(* IEC 61131-3 sources: plcassist-cli/packages/volt-lsp-iec/test-corpus/lenze-mid/Device/Plc Logic/Application/Library Manager/L_MC4P_RoboticHandling (part 2) *)

(* ---- L_MC4P_GROUPDIGITALSWITCHHANDLER.fb ---- *)
FUNCTION_BLOCK L_MC4P_GROUPDIGITALSWITCHHANDLER EXTENDS L_MC4P_Template_AG_KIN
VAR_INPUT
	XENABLE : BOOL;
	XRESETSWITCHES : BOOL;
END_VAR
VAR_OUTPUT
	XVALID : BOOL;
	XBUSY : BOOL;
	XERROR : BOOL;
	EERRORID : L_IE1P_Error;
	DWDIGITALSWITCHES : DWORD;
END_VAR
VAR
	ADWDIGITALSWITCHES : ARRAY [1..cwNbrOfdwDigSwitches] OF DWORD;
	LRPASSEDLENGTHOFSEGMENTID : LREAL;
	LRPASSEDTIMEOFSEGMENTID : LREAL;
	_MODEL : L_UBUP_BehaviourModel_LCon;
	XRESETSWITCHESOLD : BOOL;
	RSCSWITCHINGFUN : REFERENCE TO L_MC4P_SwitchingFunctionData;
	ALRSWITCHPARAMSORTED : ARRAY [1..L_MC4P_Constants.gciMaxNumParallelSwitchingFun] OF LREAL;
	XPOSRELATED : BOOL;
	ISWITCHIDXVISU : INT := 1;
	WVISUIDX : WORD := 1;
	CWNBROFDWDIGSWITCHES : WORD := 1024;
	IDXMAX : DINT;
	IDXMIN : DINT;
END_VAR
END_FUNCTION_BLOCK

METHOD ANALYZEANDSORTDATA : BOOL
VAR_INPUT
	PLISTELEMENT : POINTER TO L_MC4P_ListElement;
END_VAR
END_METHOD

METHOD GETDIGITALSWITCH : BOOL
VAR_INPUT
	WDIGITALSWITCH : WORD;
END_VAR
END_METHOD

METHOD RESET : BOOL
END_METHOD

METHOD SETDIGITALSWITCH : BOOL
VAR_INPUT
	WDIGITALSWITCH : WORD;
	XVALUE : BOOL;
END_VAR
END_METHOD

METHOD SETEVALUATEDFLAG : BOOL
VAR_INPUT
	PLISTELEMENT : POINTER TO L_MC4P_ListElement;
	IDX : INT;
END_VAR
END_METHOD

METHOD SPLITINDEX : BOOL
VAR_INPUT
	WSWITCHIDX : WORD;
END_VAR
VAR_OUTPUT
	WARRIDX : WORD;
	WBITIDX : WORD;
END_VAR
END_METHOD

METHOD CYCLICIPOCALL : BOOL
VAR_INPUT
	PLISTELEMENT : POINTER TO L_MC4P_ListElement;
	RSCCYCLICDATA : REFERENCE TO L_MC4P_CyclicData;
END_VAR
END_METHOD

METHOD FINALIZESEGMENT : BOOL
VAR_INPUT
	PLISTELEMENTACT : POINTER TO L_MC4P_ListElement;
	PLISTELEMENTNEXT : POINTER TO L_MC4P_ListElement;
END_VAR
END_METHOD

METHOD CYCLICACTION
VAR_INPUT
	ITFTIMINGCONTROLLER : L_UBUP.L_UBUP_ITimingController;
END_VAR
VAR_OUTPUT
	XCOMPLETE : BOOL;
	XABORT : BOOL;
	IERRORID : INT;
END_VAR
END_METHOD

METHOD FINALIZEACTION
VAR_INPUT
	XABORTPROPOSED : BOOL;
	IERRORIDPROPOSED : INT;
END_VAR
VAR_OUTPUT
	XCOMPLETE : BOOL;
	XABORT : BOOL;
	IERRORID : INT;
END_VAR
END_METHOD

METHOD RESETACTION
VAR_OUTPUT
	XCOMPLETE : BOOL;
END_VAR
END_METHOD

METHOD STARTACTION
VAR_OUTPUT
	XCOMPLETE : BOOL;
	IERRORID : INT;
END_VAR
END_METHOD

METHOD EXCHANGE : BOOL
VAR_INPUT
	IDX1 : DINT;
	IDX2 : DINT;
END_VAR
END_METHOD

METHOD GETVALUE : LREAL
VAR_INPUT
	IDX : DINT;
END_VAR
END_METHOD

(* ---- L_MC4P_GROUPHOME_INTERNAL.fb ---- *)
FUNCTION_BLOCK L_MC4P_GROUPHOME_INTERNAL EXTENDS L_UBUP_PoolInstance
VAR_INPUT
	EXECUTE : BOOL;
END_VAR
VAR_OUTPUT
	DONE : BOOL;
	BUSY : BOOL;
	ACTIVE : BOOL;
	COMMANDABORTED : BOOL;
	ERROR : BOOL;
	ERRORID : L_IE1P_Error;
	AXISDONE : ARRAY [1..12] OF BOOL;
END_VAR
VAR
	COORDSYSTEM : L_MC4P_CoordSystem := L_MC4P_CoordSystem.ACS;
	AMC_HOME : ARRAY [1..12] OF L_MC1P_Home_Internal;
	AMC_HOME_FBBASE : ARRAY [1..12] OF L_MC1P_Template;
	XRESETOUTPUT : BOOL;
	XEXECUTEOLD : BOOL;
	XVALIDAXISSTATES : BOOL;
	IDX : WORD;
	EACTHOMINGORDER : L_MC4P_HomingOrder := L_MC4P_HomingOrder.NoHoming;
	AXAXESHOMED : ARRAY [1..12] OF BOOL;
	ALRPOSITION_INT : ARRAY [1..12] OF LREAL;
	AEHOMINGORDER_INT : ARRAY [1..12] OF L_MC4P_HomingOrder := [12(0)];
	ECOORDSYSTEM_INT : L_MC4P_CoordSystem;
	ASCEXTPARAMETER_INT : ARRAY [1..12] OF L_MC1P_HomeParameter;
	AXUSEEXTPARAMETER_INT : ARRAY [1..12] OF BOOL;
	ASCEXTTP_INT : ARRAY [1..12] OF MC_TRIGGER_REF;
	CLASSID : DINT;
END_VAR
END_FUNCTION_BLOCK

METHOD MAIN
VAR_IN_OUT
	AXESGROUP : AXES_GROUP_KIN;
	FBBASE : L_MC4P_Template_AG_KIN;
	POSITION : ARRAY [1..12] OF LREAL;
	HOMINGORDER : ARRAY [1..12] OF L_MC4P_HomingOrder;
	HOMEABSSWITCH : ARRAY [1..12] OF BOOL;
	USEEXTPARAMETER : ARRAY [1..12] OF BOOL;
	EXTPARAMETER : ARRAY [1..12] OF L_MC1P_HomeParameter;
	EXTTP : ARRAY [1..12] OF MC_TRIGGER_REF;
END_VAR
END_METHOD

METHOD RESETOUTPUTS
END_METHOD

METHOD SETAXISMC_HOME_ACS : BOOL
VAR_IN_OUT
	AXESGROUP : AXES_GROUP_KIN;
	FBBASE : L_MC4P_Template_AG_KIN;
	HOMEABSSWITCH : ARRAY [1..12] OF BOOL;
END_VAR
END_METHOD

METHOD SETNEXTHOMESTEP
END_METHOD

METHOD GET_EERRORID : L_IE1P_Error
END_METHOD

METHOD GET_XACTIVE : BOOL
END_METHOD

METHOD GET_XBUSY : BOOL
END_METHOD

METHOD GET_XCOMMANDABORTED : BOOL
END_METHOD

METHOD GET_XDONE : BOOL
END_METHOD

METHOD GET_XINITIAL : BOOL
END_METHOD

METHOD FREE : BOOL
END_METHOD

(* ---- L_MC4P_GROUPMANUALMODE.fb ---- *)
FUNCTION_BLOCK L_MC4P_GROUPMANUALMODE EXTENDS L_MC4P_Template_AG_KIN
VAR_INPUT
	ALRSETPOSDIST : ARRAY [1..12] OF LREAL;
	SCPAR : L_MC4P_GroupManualMode_Parameter;
	ECOORDSYSTEM : L_MC4P_CoordSystem;
	AXJOGPOS : ARRAY [1..12] OF BOOL;
	AXJOGNEG : ARRAY [1..12] OF BOOL;
	AXMOVEABSEXECUTE : ARRAY [1..12] OF BOOL;
	AXMOVERELEXECUTE : ARRAY [1..12] OF BOOL;
END_VAR
VAR_OUTPUT
	XINTERNALCONTROLACTIVE : BOOL;
	XBUSY : BOOL;
	XDONE : BOOL;
	XERROR : BOOL;
	EERRORID : L_IE1P_Error;
	EMANUALMODE : L_MC4P_ManualMode := L_MC4P_ManualMode.Standby;
END_VAR
VAR
	MANMODE : L_MC4P_GroupManualMode_Internal;
END_VAR
END_FUNCTION_BLOCK

(* ---- L_MC4P_GROUPMANUALMODE_INTERNAL.fb ---- *)
FUNCTION_BLOCK L_MC4P_GROUPMANUALMODE_INTERNAL EXTENDS L_UBUP_PoolInstance
VAR_INPUT
	ALRSETPOSDIST : ARRAY [1..12] OF LREAL;
	SCPAR : L_MC4P_GroupManualMode_Parameter;
	ECOORDSYSTEM : L_MC4P_CoordSystem;
	AXJOGPOS : ARRAY [1..12] OF BOOL;
	AXJOGNEG : ARRAY [1..12] OF BOOL;
	AXMOVEABSEXECUTE : ARRAY [1..12] OF BOOL;
	AXMOVERELEXECUTE : ARRAY [1..12] OF BOOL;
	XISV2 : BOOL := FALSE;
END_VAR
VAR_OUTPUT
	XINTERNALCONTROLACTIVE : BOOL;
	XBUSY : BOOL;
	XDONE : BOOL;
	XERROR : BOOL;
	EERRORID : L_IE1P_Error;
	EMANUALMODE : L_MC4P_ManualMode := L_MC4P_ManualMode.Standby;
END_VAR
VAR
	AXMOVEABSEXECUTEEDGE : ARRAY [1..12] OF BOOL;
	AXMOVERELEXECUTEEDGE : ARRAY [1..12] OF BOOL;
	ECOORDSYSTEM_INT : L_MC4P_CoordSystem := L_MC4P_CoordSystem.MCS;
	XDOSTATEMACHINE : BOOL;
	XCHANGETOSTANDBY : BOOL := FALSE;
	XJOGGING : BOOL;
	XMOVEABSEDGE : BOOL;
	XMOVERELEDGE : BOOL;
	XMOVEABS : BOOL;
	XMOVEREL : BOOL;
	AMANUALJOG : ARRAY [1..12] OF L_MC1P_ManualJog_Internal;
	AMANUALJOG_FBBASE : ARRAY [1..12] OF L_MC1P.L_MC1P_Template;
	AMC_MOVERELATIVE : ARRAY [1..12] OF L_MC1P_MoveRelative_Internal;
	AMC_MOVERELATIVE_FBBASE : ARRAY [1..12] OF L_MC1P.L_MC1P_Template;
	AMC_MOVEABSOLUTE : ARRAY [1..12] OF L_MC1P_MoveAbsolute_Inernal;
	AMC_MOVEABSOLUTE_FBBASE : ARRAY [1..12] OF L_MC1P.L_MC1P_Template;
	EMANUALMODEOLD : L_MC4P_ManualMode := L_MC4P_ManualMode.Standby;
	ECOORDSYSTEMOLD : L_MC4P_CoordSystem;
	AXMOVEABSEXECUTEOLD : ARRAY [1..12] OF BOOL;
	AXMOVERELEXECUTEOLD : ARRAY [1..12] OF BOOL;
	XMOTIONACTIVE : BOOL := FALSE;
	APG : ARRAY [1..6] OF L_MC1P.L_MC1P_PosProfiler;
	ASCPROFILEPARAMETER : ARRAY [1..6] OF L_MC1P_ProfileParameter;
	PCOORDTRAFO : POINTER TO L_MC4P_CoordTrafo;
	COORDTRAFO_INT : L_MC4P_CoordTrafo;
	ALRPCSSETPOSATEXECUTE : ARRAY [1..6] OF LREAL;
	PLRDUMMY : POINTER TO LREAL;
	ALRPCSSETPOS_EXT : ARRAY [1..6] OF LREAL;
	ALRWCSSETPOS_EXT : ARRAY [1..6] OF LREAL;
	CLASSID : DINT;
END_VAR
END_FUNCTION_BLOCK

METHOD MAIN
VAR_IN_OUT
	AXESGROUP : AXES_GROUP_KIN;
	FBBASE : L_MC4P_Template_AG_KIN;
END_VAR
END_METHOD

METHOD GET_EERRORID : L_IE1P_Error
END_METHOD

METHOD GET_XACTIVE : BOOL
END_METHOD

METHOD GET_XBUSY : BOOL
END_METHOD

METHOD GET_XCOMMANDABORTED : BOOL
END_METHOD

METHOD GET_XDONE : BOOL
END_METHOD

METHOD GET_XINITIAL : BOOL
END_METHOD

METHOD FREE : BOOL
END_METHOD

METHOD CHECKPCSMCS : BOOL
END_METHOD

METHOD ENTRYSTANDBYSTATE
VAR_IN_OUT
	AXESGROUP : AXES_GROUP_KIN;
	FBBASE : L_MC4P_Template_AG_KIN;
END_VAR
END_METHOD

METHOD EXITMOVESTATE
VAR_IN_OUT
	AXESGROUP : AXES_GROUP_KIN;
	FBBASE : L_MC4P_Template_AG_KIN;
END_VAR
END_METHOD

METHOD GETTCSPOSINPCSMCS
VAR_INPUT
	EROTATIONCONVENTIONPCS : L_UMTP_RotationConvention;
END_VAR
VAR_IN_OUT
	AXESGROUP : AXES_GROUP_KIN;
	ALRPCSSETPOS : ARRAY [1..6] OF LREAL;
END_VAR
END_METHOD

METHOD ISMOTIONALLOWED
VAR_IN_OUT
	AXESGROUP : AXES_GROUP_KIN;
	FBBASE : L_MC4P_Template_AG_KIN;
	SCPAR : L_MC4P_GroupManualMode_Parameter;
	ECOORDSYSTEM : L_MC4P_CoordSystem;
	AXJOGPOS : ARRAY [1..12] OF BOOL;
	AXJOGNEG : ARRAY [1..12] OF BOOL;
	AXMOVEABSEXECUTE : ARRAY [1..12] OF BOOL;
	AXMOVERELEXECUTE : ARRAY [1..12] OF BOOL;
END_VAR
END_METHOD

METHOD JOGAXISREF
VAR_INPUT
	XWCS : BOOL;
	XACS : BOOL;
	XAUX : BOOL;
END_VAR
VAR_IN_OUT
	AXESGROUP : AXES_GROUP_KIN;
	FBBASE : L_MC4P_Template_AG_KIN;
	SCPAR : L_MC4P_GroupManualMode_Parameter;
	AXJOGPOS : ARRAY [1..12] OF BOOL;
	AXJOGNEG : ARRAY [1..12] OF BOOL;
END_VAR
END_METHOD

METHOD JOGPCSMCS
VAR_IN_OUT
	AXESGROUP : AXES_GROUP_KIN;
	FBBASE : L_MC4P_Template_AG_KIN;
	SCPAR : L_MC4P_GroupManualMode_Parameter;
	AXJOGPOS : ARRAY [1..12] OF BOOL;
	AXJOGNEG : ARRAY [1..12] OF BOOL;
END_VAR
END_METHOD

METHOD MOVEABSAXISREF
VAR_INPUT
	XWCS : BOOL;
	XACS : BOOL;
	XAUX : BOOL;
END_VAR
VAR_IN_OUT
	AXESGROUP : AXES_GROUP_KIN;
	FBBASE : L_MC4P_Template_AG_KIN;
	ALRSETPOSDIST : ARRAY [1..12] OF LREAL;
	SCPAR : L_MC4P_GroupManualMode_Parameter;
	AXMOVEABSEXECUTE : ARRAY [1..12] OF BOOL;
END_VAR
END_METHOD

METHOD MOVEABSPCSMCS
VAR_IN_OUT
	AXESGROUP : AXES_GROUP_KIN;
	FBBASE : L_MC4P_Template_AG_KIN;
	ALRSETPOSDIST : ARRAY [1..12] OF LREAL;
	SCPAR : L_MC4P_GroupManualMode_Parameter;
	AXMOVEABSEXECUTE : ARRAY [1..12] OF BOOL;
END_VAR
END_METHOD

METHOD MOVERELAXISREF
VAR_INPUT
	XWCS : BOOL;
	XACS : BOOL;
	XAUX : BOOL;
END_VAR
VAR_IN_OUT
	AXESGROUP : AXES_GROUP_KIN;
	FBBASE : L_MC4P_Template_AG_KIN;
	ALRSETPOSDIST : ARRAY [1..12] OF LREAL;
	SCPAR : L_MC4P_GroupManualMode_Parameter;
	AXMOVERELEXECUTE : ARRAY [1..12] OF BOOL;
END_VAR
END_METHOD

METHOD MOVERELPCSMCS
VAR_IN_OUT
	AXESGROUP : AXES_GROUP_KIN;
	FBBASE : L_MC4P_Template_AG_KIN;
	ALRSETPOSDIST : ARRAY [1..12] OF LREAL;
	SCPAR : L_MC4P_GroupManualMode_Parameter;
	AXMOVERELEXECUTE : ARRAY [1..12] OF BOOL;
END_VAR
END_METHOD

METHOD RESETMOTIONQUERY
END_METHOD

METHOD WRITEPCSMCSPOS2AXES
VAR_INPUT
	EROTATIONCONVENTIONPCS : L_UMTP_RotationConvention;
	XRELATIVE : BOOL;
END_VAR
VAR_IN_OUT
	AXESGROUP : AXES_GROUP_KIN;
	FBBASE : L_MC4P_Template_AG_KIN;
	ALRPCSSETPOS : ARRAY [1..6] OF LREAL;
	ALRPCSSETVEL : ARRAY [1..6] OF LREAL;
END_VAR
END_METHOD

METHOD CALL_AXISREFPARM
VAR_INPUT
	AXESGROUP : REFERENCE TO AXES_GROUP_KIN;
	LRVELOCITY : REFERENCE TO LREAL;
	LRACCELERATION : REFERENCE TO LREAL;
	LRDECELERATION : REFERENCE TO LREAL;
	LRJERK : REFERENCE TO LREAL;
	AXIS_IDX_LOCAL : WORD;
END_VAR
END_METHOD

METHOD CALL_PCSMCSPARM
VAR_INPUT
	AXESGROUP : REFERENCE TO AXES_GROUP_KIN;
	ALRPCSSETPOS : REFERENCE TO ARRAY [1..6] OF LREAL;
	IDX_LOCAL : WORD;
END_VAR
END_METHOD

(* ---- L_MC4P_GROUPPOWER.fb ---- *)
FUNCTION_BLOCK L_MC4P_GROUPPOWER EXTENDS L_MC4P_Template_AG_REF
VAR_INPUT
	XENABLE : BOOL;
	AEAXISENABLE : ARRAY [1..12] OF L_MC4P_AxisEnableMode := [12(L_MC4P_AxisEnableMode.EnablePosNeg)];
END_VAR
VAR_OUTPUT
	XSTATUS : BOOL;
	XVALID : BOOL;
	XERROR : BOOL;
	EERRORID : L_IE1P_Error;
END_VAR
VAR
	AMC_POWER : ARRAY [1..12] OF MC_Power;
	XENABLEOLD : BOOL;
	IDX : WORD;
	IDX_PLUSSIX : WORD;
	XAXISEXTENABLED : BOOL := FALSE;
	XERRORINTERN : BOOL := FALSE;
	EERRORIDINTERN : L_IE1P_Error;
	XAXISERROR : BOOL := FALSE;
END_VAR
END_FUNCTION_BLOCK

(* ---- L_MC4P_GROUPREADACTUALPOSITION_INTERNAL.fb ---- *)
FUNCTION_BLOCK L_MC4P_GROUPREADACTUALPOSITION_INTERNAL EXTENDS L_UBUP_Instance
VAR_INPUT
	ENABLE : BOOL;
	COORDSYSTEM : L_MC4P_CoordSystem;
END_VAR
VAR_OUTPUT
	VALID : BOOL;
	BUSY : BOOL;
	ERROR : BOOL;
	ERRORID : L_IE1P_Error;
END_VAR
VAR
	IDX : WORD;
	XENABLEOLD : BOOL;
	PCOORDTRAFO : POINTER TO L_MC4P_CoordTrafo;
	ALRPOSITIONTMP : ARRAY [1..6] OF LREAL;
	CLASSID : DINT;
END_VAR
END_FUNCTION_BLOCK

METHOD MAIN
VAR_INPUT
	XUSESETVALUES : BOOL;
END_VAR
VAR_IN_OUT
	AXESGROUP : AXES_GROUP_KIN;
	FBBASE : L_MC4P_Template_AG_KIN;
	POSITION : ARRAY [1..12] OF LREAL;
END_VAR
END_METHOD

(* ---- L_MC4P_GROUPREADACTUALVELOCITY_INTERNAL.fb ---- *)
FUNCTION_BLOCK L_MC4P_GROUPREADACTUALVELOCITY_INTERNAL EXTENDS L_UBUP_Instance
VAR_INPUT
	ENABLE : BOOL;
	COORDSYSTEM : L_MC4P_CoordSystem;
END_VAR
VAR_OUTPUT
	VALID : BOOL;
	BUSY : BOOL;
	ERROR : BOOL;
	ERRORID : L_IE1P_Error;
END_VAR
VAR
	IDX : WORD;
	XENABLEOLD : BOOL;
	ALRVELOCITYTMP1 : ARRAY [1..6] OF LREAL;
	ALRVELOCITYTMP2 : ARRAY [1..6] OF LREAL;
	ALRPOSITIONTMP : ARRAY [1..6] OF LREAL;
	PCOORDTRAFO : POINTER TO L_MC4P_CoordTrafo;
	ALRPOSVEKPCS2TCS : ARRAY [1..3] OF LREAL;
	ROT_MAT : ARRAY [1..3, 1..3] OF LREAL;
	T4 : LREAL;
	T5 : LREAL;
	T7 : LREAL;
	CLASSID : DINT;
END_VAR
END_FUNCTION_BLOCK

METHOD MAIN
VAR_INPUT
	XUSESETVALUES : BOOL;
END_VAR
VAR_IN_OUT
	AXESGROUP : AXES_GROUP_KIN;
	FBBASE : L_MC4P_Template_AG_KIN;
	VELOCITY : ARRAY [1..12] OF LREAL;
	PATHVELOCITY : LREAL;
END_VAR
END_METHOD

(* ---- L_MC4P_GROUPREADSTATUS_INTERNAL.fb ---- *)
FUNCTION_BLOCK L_MC4P_GROUPREADSTATUS_INTERNAL EXTENDS L_UBUP_PoolInstance
VAR_INPUT
	ENABLE : BOOL;
END_VAR
VAR_OUTPUT
	VALID : BOOL;
	BUSY : BOOL;
	ERROR : BOOL;
	ERRORID : L_IE1P_Error;
	GROUPMOVING : BOOL;
	GROUPHOMING : BOOL;
	GROUPERRORSTOP : BOOL;
	GROUPSTANDBY : BOOL;
	GROUPSTOPPING : BOOL;
	GROUPDISABLED : BOOL;
	CONSTANTVELOCITY : BOOL;
	ACCELERATING : BOOL;
	DECELERATING : BOOL;
	INPOSITION : BOOL;
	STANDSTILL : BOOL;
END_VAR
VAR
	XENABLEOLD : BOOL;
	IDX : INT;
	CLASSID : DINT;
END_VAR
END_FUNCTION_BLOCK

METHOD MAIN
VAR_IN_OUT
	AXESGROUP : AXES_GROUP_KIN;
	FBBASE : L_MC4P_Template_AG_KIN;
END_VAR
END_METHOD

(* ---- L_MC4P_GROUPRESET_INTERNAL.fb ---- *)
FUNCTION_BLOCK L_MC4P_GROUPRESET_INTERNAL EXTENDS L_UBUP_Instance
VAR_INPUT
	EXECUTE : BOOL;
END_VAR
VAR_OUTPUT
	DONE : BOOL;
	BUSY : BOOL;
	ERROR : BOOL;
	ERRORID : L_IE1P_Error;
END_VAR
VAR
	ARESET : ARRAY [1..18] OF MC_Reset;
	PAXESGROUP : POINTER TO AXES_GROUP_KIN;
	XEXECUTEOLD : BOOL;
	PWTMP : POINTER TO WORD;
	IDX : INT;
	XRESETPOSSIBLE : BOOL;
	XRESETOUTPUT : BOOL;
	DWRESETCYCLECOUNTERSTART : DWORD;
	XNOERRORACTIVE : BOOL;
	XERRORSTOPDONE : BOOL;
	XAXESGROUPINERROR : BOOL;
	XAXISINERROR : BOOL;
	XWAITFORRESETEVENT : BOOL;
	DWMAXTIMEOUT : DWORD;
	CLASSID : DINT;
END_VAR
END_FUNCTION_BLOCK

METHOD MAIN
VAR_IN_OUT
	AXESGROUP : AXES_GROUP_REF;
	FBBASE : L_MC4P_Template_ForAG;
END_VAR
END_METHOD

METHOD REQUESTINTERFACE : BOOL
VAR_INPUT
	ID : DINT;
	PITFUNKNOWN : POINTER TO L_UBUP_IUnknown;
END_VAR
END_METHOD

(* ---- L_MC4P_GROUPSETOVERRIDE.fb ---- *)
FUNCTION_BLOCK L_MC4P_GROUPSETOVERRIDE EXTENDS L_MC4P_Template_AG_KIN
VAR_INPUT
	XENABLE : BOOL;
	LROVERRIDE : LREAL := 1.0;
	LRFADINGTIME : LREAL := 2.5;
END_VAR
VAR_OUTPUT
	XENABLED : BOOL;
	XBUSY : BOOL;
	XERROR : BOOL;
	EERRORID : L_IE1P_Error := L_IE1P_Error.NoError;
END_VAR
VAR
	GROUPSETOVERRIDE : L_MC4P_GroupSetOverride_Internal;
END_VAR
END_FUNCTION_BLOCK

(* ---- L_MC4P_GROUPSETOVERRIDE_INTERNAL.fb ---- *)
FUNCTION_BLOCK L_MC4P_GROUPSETOVERRIDE_INTERNAL EXTENDS L_UBUP_PoolInstance
VAR_INPUT
	XENABLE : BOOL;
	LROVERRIDE : LREAL := 1.0;
	LRFADINGTIME : LREAL := 2.5;
END_VAR
VAR_OUTPUT
	XENABLED : BOOL;
	XBUSY : BOOL;
	XERROR : BOOL;
	EERRORID : L_IE1P_Error := L_IE1P_Error.NoError;
END_VAR
VAR
	XENABLEOLD : BOOL;
	CLASSID : DINT;
END_VAR
END_FUNCTION_BLOCK

METHOD MAIN
VAR_IN_OUT
	AXESGROUP : AXES_GROUP_KIN;
	FBBASE : L_MC4P_Template_AG_KIN;
END_VAR
END_METHOD

METHOD REQUESTINTERFACE : BOOL
VAR_INPUT
	ID : DINT;
	PITFUNKNOWN : POINTER TO L_UBUP_IUnknown;
END_VAR
END_METHOD

(* ---- L_MC4P_GROUPSETPOSITION_INTERNAL.fb ---- *)
FUNCTION_BLOCK L_MC4P_GROUPSETPOSITION_INTERNAL EXTENDS L_UBUP_PoolInstance
VAR_INPUT
	EXECUTE : BOOL;
	RELATIVE : BOOL := FALSE;
END_VAR
VAR_OUTPUT
	DONE : BOOL;
	BUSY : BOOL;
	ACTIVE : BOOL;
	ERROR : BOOL;
	ERRORID : L_IE1P_Error;
END_VAR
VAR
	COORDSYSTEM : L_MC4P_CoordSystem := L_MC4P_CoordSystem.ACS;
	XRESETOUTPUT : BOOL;
	AMC_SETPOSITION : ARRAY [1..12] OF L_MC1P.MC_SetPosition;
	IDX : WORD;
	XEXECUTEOLD : BOOL;
	CLASSID : DINT;
END_VAR
END_FUNCTION_BLOCK

METHOD MAIN
VAR_IN_OUT
	AXESGROUP : AXES_GROUP_KIN;
	FBBASE : L_MC4P_Template_AG_KIN;
	POSITION : ARRAY [1..12] OF LREAL;
END_VAR
END_METHOD

METHOD REQUESTINTERFACE : BOOL
VAR_INPUT
	ID : DINT;
	PITFUNKNOWN : POINTER TO L_UBUP_IUnknown;
END_VAR
END_METHOD

(* ---- L_MC4P_GROUPSTOP_INTERNAL.fb ---- *)
FUNCTION_BLOCK L_MC4P_GROUPSTOP_INTERNAL EXTENDS L_MC4P_CalcStopProfiles
VAR_INPUT
	EXECUTE : BOOL;
	DECELERATION : LREAL;
	JERK : LREAL;
END_VAR
VAR_OUTPUT
	DONE : BOOL;
	BUSY : BOOL;
	ACTIVE : BOOL;
	COMMANDABORTED : BOOL;
	ERROR : BOOL;
	ERRORID : L_IE1P_Error;
END_VAR
VAR
	_ITFOWNER : L_UBUP.L_UBUP_IFBPool;
	_XWHANDLE : __XWORD;
	_XOCCUPIED : BOOL;
	LRINPUTJERK : LREAL;
	LRINPUTDECELERATION : LREAL;
	AMC_STOP : ARRAY [1..18] OF L_MC1P.L_MC1P_Stop_Internal;
	AMC_STOP_FBBASE : ARRAY [1..18] OF L_MC1P.L_MC1P_Template;
	IDX : WORD;
	XEXECUTEOLD : BOOL;
	XRESETOUTPUT : BOOL;
	XDONEINTERN : BOOL;
	XDONEOLD : BOOL;
	XERRORINTERN : BOOL;
	EERRORIDINTERN : L_IE1P_Error;
	DWINTERNALID : DWORD;
	XSTOPPROFILESCALCULATED : BOOL;
	_DWOBJID : DWORD;
	CLASSID : DINT;
	INSTANCEPTR : POINTER TO BYTE;
	OBJECTID : DWORD;
	OCCUPIED : BOOL;
END_VAR
END_FUNCTION_BLOCK

METHOD GROUPSTOPACS
VAR_IN_OUT
	AXESGROUP : AXES_GROUP_KIN;
	FBBASE : L_MC4P_Template_AG_KIN;
END_VAR
END_METHOD

METHOD GROUPSTOPMCS
VAR_IN_OUT
	AXESGROUP : AXES_GROUP_KIN;
	FBBASE : L_MC4P_Template_AG_KIN;
END_VAR
END_METHOD

METHOD MAIN
VAR_IN_OUT
	AXESGROUP : AXES_GROUP_KIN;
	FBBASE : L_MC4P_Template_AG_KIN;
END_VAR
END_METHOD

METHOD RESETOUTPUTS
VAR_IN_OUT
	AXESGROUP : AXES_GROUP_KIN;
END_VAR
END_METHOD

METHOD GET_EERRORID : L_IE1P_Error
END_METHOD

METHOD GET_XACTIVE : BOOL
END_METHOD

METHOD GET_XBUSY : BOOL
END_METHOD

METHOD GET_XCOMMANDABORTED : BOOL
END_METHOD

METHOD GET_XDONE : BOOL
END_METHOD

METHOD GET_XINITIAL : BOOL
END_METHOD

METHOD FREE : BOOL
END_METHOD

METHOD OCCUPY : BOOL
VAR_INPUT
	ITFOWNER : L_UBUP.L_UBUP_IFBPool;
	XWHANDLE : __XWORD;
END_VAR
END_METHOD

METHOD REQUESTINTERFACE : BOOL
VAR_INPUT
	ID : DINT;
	PITFUNKNOWN : POINTER TO L_UBUP_IUnknown;
END_VAR
END_METHOD

METHOD FB_INIT : BOOL
VAR_INPUT
	BINITRETAINS : BOOL;
	BINCOPYCODE : BOOL;
END_VAR
END_METHOD

(* ---- L_MC4P_GROUPTORQUEPRECONTROL.fb ---- *)
FUNCTION_BLOCK L_MC4P_GROUPTORQUEPRECONTROL EXTENDS L_MC4P_Template_AG_KIN
VAR_INPUT
	XENABLE : BOOL;
	XUSEAXESGROUPPARAM : BOOL := FALSE;
	XWRITETOPARAMETER : BOOL := FALSE;
	LRTORQUEOVERRIDE : LREAL := 0;
	LRTORQUELIMITFACTOR : LREAL := 1;
	ALRTORQUERATELIMIT : ARRAY [1..6] OF LREAL := [6(0.0)];
	LRLOADMASS : LREAL;
	ITFDYNAMICPAR : L_MC4P_DynamicPar;
END_VAR
VAR_OUTPUT
	XVALID : BOOL;
	XBUSY : BOOL;
	XERROR : BOOL;
	EERRORID : L_IE1P_Error;
	ALRSETTORQUEOUT : ARRAY [1..6] OF LREAL;
	ALRACTTORQUE : ARRAY [1..6] OF LREAL;
END_VAR
VAR
	LICHANDLING : L_IMHP_LLMHandling;
	IDX : INT;
	IDX2 : WORD;
	XENABLEOLD : BOOL;
	XWRITETOPARAMETEROLD : BOOL;
	ALRTORQUELIMITS : ARRAY [1..6] OF LREAL;
	ALRTORQUEDELTACYCLE : ARRAY [1..6] OF LREAL := [6(0.0)];
	XUSEFILTEREDVALUES : BOOL := TRUE;
	XSETVALUEFILTERACTIVE : BOOL;
	EBEHAVEONERRORSTOP : L_MC4P_ErrorStopBehaviour := L_MC4P_ErrorStopBehaviour.SetTorqueToZero;
	ALRGRAVITATION : ARRAY [1..3] OF LREAL;
	ALRCOULOMBFRIC : ARRAY [1..6] OF LREAL;
	ALRVISCFRIC : ARRAY [1..6] OF LREAL;
	ALRDYNAMICPAR : ARRAY [1..L_MC4P_Constants.uimaxNbrOfDynamicPar] OF LREAL;
	EERRORTMP : L_IE1P_Error;
	ALRTOOLINERTIA : ARRAY [1..3, 1..3] OF LREAL;
	ALRLOADINERTIA : ARRAY [1..3, 1..3] OF LREAL;
	BEHAVEONERRORSTOP : L_MC4P_ErrorStopBehaviour;
	USEFILTEREDVALUES : BOOL;
END_VAR
END_FUNCTION_BLOCK

(* ---- L_MC4P_GROUPWAITTIME.fb ---- *)
FUNCTION_BLOCK L_MC4P_GROUPWAITTIME EXTENDS L_MC4P_Template_MoveLicence
VAR_INPUT
	XEXECUTE : BOOL;
	LRTIME : LREAL;
END_VAR
VAR_OUTPUT
	XDONE : BOOL;
	XBUSY : BOOL;
	XACTIVE : BOOL;
	XCOMMANDABORTED : BOOL;
	XERROR : BOOL;
	EERRORID : L_IE1P_Error;
END_VAR
VAR
	WAIT : L_MC4P_GroupWaitTime_Internal;
	PMOVE : POINTER TO L_MC4P_MoveContPath;
END_VAR
END_FUNCTION_BLOCK

(* ---- L_MC4P_GROUPWAITTIME_INTERNAL.fb ---- *)
FUNCTION_BLOCK L_MC4P_GROUPWAITTIME_INTERNAL EXTENDS L_MC4P_MoveContPath
VAR_INPUT
	XEXECUTE : BOOL;
	LRTIME : LREAL;
END_VAR
VAR_OUTPUT
	XDONE : BOOL;
	XBUSY : BOOL;
	XACTIVE : BOOL;
	XCOMMANDABORTED : BOOL;
	XERROR : BOOL;
	EERRORID : L_IE1P_Error;
END_VAR
VAR
	LRTIME_INPUT : LREAL;
	AEAUXMODE : ARRAY [1..6] OF L_MC4P_AuxMode := [6(L_MC4P_AuxMode.Inactive)];
	TRANSITIONPARAMETER : ARRAY [1..12] OF LREAL := [12(0)];
	COORDSYSTEM : L_MC4P_CoordSystem;
	BUFFERMODE : MC_BUFFER_MODE;
	TRANSITIONMODE : MC_TRANSITION_MODE;
	CLASSID : DINT;
END_VAR
END_FUNCTION_BLOCK

METHOD HOMINGREQUIRED : BOOL
END_METHOD

METHOD ISPTP : BOOL
END_METHOD

METHOD MAIN
VAR_IN_OUT
	AXESGROUP : AXES_GROUP_KIN;
	FBBASE : L_MC4P_Template_AG_KIN;
END_VAR
END_METHOD

METHOD PARAMETERFREEZE
VAR_IN_OUT
	AXESGROUP : AXES_GROUP_KIN;
	FBBASE : L_MC4P_Template_AG_KIN;
	COORDSYSTEM : L_MC4P_CoordSystem;
	BUFFERMODE : MC_BUFFER_MODE;
	TRANSITIONMODE : MC_TRANSITION_MODE;
	TRANSITIONPARAMETER : ARRAY [1..12] OF LREAL;
END_VAR
END_METHOD

METHOD SETPATHELEMENT
VAR_IN_OUT
	AXESGROUP : AXES_GROUP_KIN;
	FBBASE : L_MC4P_Template_AG_KIN;
	ALRSTARTPOS : ARRAY [1..12] OF LREAL;
	ALRSUPERPOSPOSATSTART : ARRAY [1..3] OF LREAL;
END_VAR
END_METHOD

(* ---- L_MC4P_INTERPOLATEPATH.fb ---- *)
FUNCTION_BLOCK L_MC4P_INTERPOLATEPATH
VAR_INPUT
	PLIST : POINTER TO L_MC4P_PathDataList;
	PAXESGROUP : POINTER TO AXES_GROUP_KIN;
	XEXCLUDEAUX : BOOL := FALSE;
	XIGNOREOVERRIDEWAITTIME : BOOL := FALSE;
	ITFDIGSWITCHOBSERVER : L_MC4P_IDigSwitchHandling;
END_VAR
VAR_OUTPUT
	AXAUXAXISACTIVE : ARRAY [1..6] OF BOOL;
	NSEGMENTNO : DINT;
	XERROR : BOOL := FALSE;
	EERRORID : L_IE1P_Error;
	DWINTERNALID : DWORD;
END_VAR
VAR
	SCCYCLICDATA : L_MC4P_CyclicData;
	PLISTELEMENTTIME : POINTER TO L_MC4P_ListElement;
	PLISTELEMENTGEO : POINTER TO L_MC4P_ListElement;
	PLISTELEMENTTOBODELETED : POINTER TO L_MC4P_ListElement;
	XREADY : BOOL;
	PATHFILTER : L_MC4P_SetValueFilter;
	AROTFILTER : ARRAY [1..3] OF L_MC4P_SetValueFilter;
	AAUXFILTER : ARRAY [1..6] OF L_MC4P_SetValueFilter;
	EFILTERMODE : L_MC4P_SetValueFilterMode := L_MC4P_SetValueFilterMode.EqualySpaced;
	UIFILTERTIME : UINT;
	XENABLEFILTER : BOOL;
	XAXESGROUPIPOSTANDSTILL : BOOL := TRUE;
	PPAUSEDTIMEELEMENT : POINTER TO L_MC4P_ListElement;
	XPAUSETIMEIPO : BOOL;
	XRELEASETIMEIPO : BOOL;
	AXAUXAXISACTIVEOLD : ARRAY [1..6] OF BOOL;
	XFIRSTCALLOFNEWSEQUENCE : BOOL;
END_VAR
END_FUNCTION_BLOCK

METHOD AXISPASSEDTARGETPOS : BOOL
VAR_INPUT
	ETRAVERSINGRANGE : L_MC1P_TraversingRange;
	LRCYCLELENGTH : LREAL;
	LRSTARTPOS : LREAL;
	LRTARGETPOS : LREAL;
	LRIPOPOS : LREAL;
	LRIPOVEL : LREAL;
	LRIPOACC : LREAL;
	LRIPOPOSOLD : LREAL;
	SCPROFILEDATAACT : REFERENCE TO L_MC1P_ProfileData;
	SCPROFILEDATANEXT : REFERENCE TO L_MC1P_ProfileData;
END_VAR
END_METHOD

METHOD ENDSWITHRESTPHASE : BOOL
VAR_IN_OUT
	PROFILEDATA : L_MC1P_ProfileData;
END_VAR
END_METHOD

METHOD GEOMETRYPASSED : BOOL
VAR_IN_OUT
	PLISTELEMENT : POINTER TO L_MC4P_ListElement;
	SCCYCLICDATA : L_MC4P_CyclicData;
END_VAR
END_METHOD

METHOD GETSTARTDIRECTION : MC_Direction
VAR_IN_OUT
	PROFILEDATA : L_MC1P_ProfileData;
END_VAR
END_METHOD

METHOD GETTARGETDIRECTION : MC_Direction
VAR_IN_OUT
	PROFILEDATA : L_MC1P_ProfileData;
END_VAR
END_METHOD

METHOD INITIPO
END_METHOD

METHOD INTERPOLATECPGEOMETRY
VAR_IN_OUT
	PLISTELEMENTGEO : POINTER TO L_MC4P_ListElement;
	SCCYCLICDATA : L_MC4P_CyclicData;
END_VAR
END_METHOD

METHOD INTERPOLATETIMEPROFILES
VAR_IN_OUT
	PLISTELEMENTTIME : POINTER TO L_MC4P_ListElement;
	SCCYCLICDATA : L_MC4P_CyclicData;
END_VAR
END_METHOD

METHOD INTERPOLATOR
VAR_IN_OUT
	PLISTELEMENTTIME : POINTER TO L_MC4P_ListElement;
	PLISTELEMENTGEO : POINTER TO L_MC4P_ListElement;
	SCCYCLICDATA : L_MC4P_CyclicData;
END_VAR
END_METHOD

METHOD ISCARTESIAN : BOOL
VAR_INPUT
	ESEGMENTTYPE : L_MC4P_SegmentType;
END_VAR
END_METHOD

METHOD MODULOFILTEROVERRIDE
VAR_IN_OUT
	PLISTELEMENTTIME : POINTER TO L_MC4P_ListElement;
	SCCYCLICDATA : L_MC4P_CyclicData;
END_VAR
END_METHOD

METHOD RESETIPO
END_METHOD

METHOD TARGETVELOFLISTELEMENTEQ0 : BOOL
VAR_INPUT
	PLISTELEMENT : POINTER TO L_MC4P_ListElement;
END_VAR
END_METHOD

(* ---- L_MC4P_KIN_REF_GENERIC.fb ---- *)
FUNCTION_BLOCK L_MC4P_KIN_REF_GENERIC
VAR_OUTPUT
	XACTIVE : BOOL;
END_VAR
VAR
	PAXESGROUP : POINTER TO Axes_Group_KIN;
END_VAR
END_FUNCTION_BLOCK

METHOD GETPARAITF : L_MC4P_IKinParamExtern
END_METHOD

METHOD GETTRAFOITF : L_MC4P_ITrafoExtern
END_METHOD

METHOD LINKEDAXESGROUP_GET : POINTER TO AXES_GROUP_KIN
END_METHOD

METHOD LINKEDAXESGROUP_SET
VAR_INPUT
	LINKEDAXESGROUP : POINTER TO AXES_GROUP_KIN;
END_VAR
END_METHOD

METHOD SETACSAXISTYPE
VAR_OUTPUT
	AEAXES : ARRAY [1..6] OF L_MC4P_AxisType := [L_MC4P_AxisType.linear, L_MC4P_AxisType.linear, L_MC4P_AxisType.linear, L_MC4P_AxisType.rotary, L_MC4P_AxisType.unconnected, L_MC4P_AxisType.unconnected];
END_VAR
END_METHOD

METHOD SETINITIALVALUESOFCONSTANTMCSAXES
VAR_OUTPUT
	ALRMCSPOS : ARRAY [1..6] OF LREAL := [0.0, 0.0, 0.0, 180.0, 0.0, 0.0];
END_VAR
END_METHOD

METHOD SETMCSAXISTYPE
VAR_OUTPUT
	AEAXES : ARRAY [1..6] OF L_MC4P_AxisType := [L_MC4P_AxisType.linear, L_MC4P_AxisType.linear, L_MC4P_AxisType.linear, L_MC4P_AxisType.unconnected, L_MC4P_AxisType.unconnected, L_MC4P_AxisType.rotary];
END_VAR
END_METHOD

METHOD CALCULATEPARAMETER
END_METHOD

METHOD CHECKPARAMETER : BOOL
END_METHOD

METHOD PARAMETERCHANGED
END_METHOD

METHOD CALCBACKWARDTRAFO : WORD
VAR_IN_OUT
	AXESGROUP : AXES_GROUP_KIN;
	ALRPOSFLANGE : ARRAY [1..6] OF LREAL;
	ALRPOSAXES : ARRAY [1..6] OF LREAL;
	AICONFIGURATION : ARRAY [1..6] OF INT;
END_VAR
END_METHOD

METHOD CALCFORWARDTRAFO : WORD
VAR_IN_OUT
	AXESGROUP : AXES_GROUP_KIN;
	ALRPOSFLANGE : ARRAY [1..6] OF LREAL;
	ALRPOSAXES : ARRAY [1..6] OF LREAL;
END_VAR
END_METHOD

METHOD CALCULATECONFIGURATION : WORD
VAR_IN_OUT
	AXESGROUP : AXES_GROUP_KIN;
	ALRPOSFLANGE : ARRAY [1..6] OF LREAL;
	ALRPOSAXES : ARRAY [1..6] OF LREAL;
	AICONFIGURATION : ARRAY [1..6] OF INT;
END_VAR
END_METHOD

(* ---- L_MC4P_KINCOORDPROVIDER.fb ---- *)
FUNCTION_BLOCK L_MC4P_KINCOORDPROVIDER
VAR_INPUT
	ALRACSPOS : ARRAY [1..6] OF LREAL;
	ALRACSVEL : ARRAY [1..6] OF LREAL;
	ALRACSACC : ARRAY [1..6] OF LREAL;
	ALRJCSPOS : ARRAY [1..6] OF LREAL;
	ALRJCSVEL : ARRAY [1..6] OF LREAL;
	ALRJCSACC : ARRAY [1..6] OF LREAL;
	ALRFCSPOS : ARRAY [1..6] OF LREAL;
	ALRFCSVEL : ARRAY [1..6] OF LREAL;
	ALRFCSACC : ARRAY [1..6] OF LREAL;
	ALRMCSPOS : ARRAY [1..6] OF LREAL;
	ALRMCSVEL : ARRAY [1..6] OF LREAL;
	ALRMCSACC : ARRAY [1..6] OF LREAL;
	ALRWCSPOS : ARRAY [1..6] OF LREAL;
	ALRWCSVEL : ARRAY [1..6] OF LREAL;
	ALRWCSACC : ARRAY [1..6] OF LREAL;
	SCFCSFRAME : L_UMTP_RobotFrame;
	SCMCSFRAME : L_UMTP_RobotFrame;
	SCWCSFRAME : L_UMTP_RobotFrame;
END_VAR
VAR_OUTPUT
	UDILOWERSYSTEM : UDINT := 0;
	UDIUPPERSYSTEM : UDINT := 0;
	UDIDIM : UDINT := 0;
	PLRACSPOS : POINTER TO LREAL;
	PLRACSVEL : POINTER TO LREAL;
	PLRACSACC : POINTER TO LREAL;
	PLRJCSPOS : POINTER TO LREAL;
	PLRJCSVEL : POINTER TO LREAL;
	PLRJCSACC : POINTER TO LREAL;
	PLRFCSPOS : POINTER TO LREAL;
	PLRFCSVEL : POINTER TO LREAL;
	PLRFCSACC : POINTER TO LREAL;
	PLRMCSPOS : POINTER TO LREAL;
	PLRMCSVEL : POINTER TO LREAL;
	PLRMCSACC : POINTER TO LREAL;
	PLRWCSPOS : POINTER TO LREAL;
	PLRWCSVEL : POINTER TO LREAL;
	PLRWCSACC : POINTER TO LREAL;
	PFCSFRAME : POINTER TO L_UMTP_RobotFrame;
	PMCSFRAME : POINTER TO L_UMTP_RobotFrame;
	PWCSFRAME : POINTER TO L_UMTP_RobotFrame;
END_VAR
VAR
	ACSACC : POINTER TO LREAL;
	ACSPOS : POINTER TO LREAL;
	ACSVEL : POINTER TO LREAL;
	DIM : UDINT;
	FCSACC : POINTER TO LREAL;
	FCSFRAME : POINTER TO L_UMTP_RobotFrame;
	FCSPOS : POINTER TO LREAL;
	FCSVEL : POINTER TO LREAL;
	JCSACC : POINTER TO LREAL;
	JCSPOS : POINTER TO LREAL;
	JCSVEL : POINTER TO LREAL;
	LOWERSYSTEM : UDINT;
	MCSACC : POINTER TO LREAL;
	MCSFRAME : POINTER TO L_UMTP_RobotFrame;
	MCSPOS : POINTER TO LREAL;
	MCSVEL : POINTER TO LREAL;
	UPPERSYSTEM : UDINT;
	WCSACC : POINTER TO LREAL;
	WCSFRAME : POINTER TO L_UMTP_RobotFrame;
	WCSPOS : POINTER TO LREAL;
	WCSVEL : POINTER TO LREAL;
END_VAR
END_FUNCTION_BLOCK

METHOD EQUALS : BOOL
VAR_INPUT
	ITFPROVIDER : L_MC4P_IKinCoordProvider;
	UDISYSTEM : UDINT;
	XPOS : BOOL;
	XVEL : BOOL;
	XACC : BOOL;
END_VAR
END_METHOD

METHOD FB_INIT : BOOL
VAR_INPUT
	BINITRETAINS : BOOL;
	BINCOPYCODE : BOOL;
END_VAR
END_METHOD

METHOD FB_REINIT : BOOL
END_METHOD

METHOD COPYFRAME
VAR_INPUT
	PSCFRAME : POINTER TO L_UMTP_RobotFrame;
END_VAR
VAR_IN_OUT
	SCFRAME : L_UMTP_RobotFrame;
END_VAR
END_METHOD

METHOD COPYVECTOR
VAR_INPUT
	PLR : POINTER TO LREAL;
END_VAR
VAR_IN_OUT
	ALR : ARRAY [1..6] OF LREAL;
END_VAR
END_METHOD

METHOD CLEAR
END_METHOD

METHOD COPYFROM
VAR_INPUT
	ICOORD : L_MC4P_IKinCoordProvider;
	ELEVEL : INT;
END_VAR
END_METHOD

METHOD SETDIM
VAR_INPUT
	UDIDIM : UDINT;
END_VAR
END_METHOD

METHOD SETLOWERSYSTEM
VAR_INPUT
	UDILOWER : UDINT;
END_VAR
END_METHOD

METHOD SETUPPERSYSTEM
VAR_INPUT
	UDIUPPER : UDINT;
END_VAR
END_METHOD

METHOD THRESHOLD
VAR_INPUT
	LRTHRESHOLD : LREAL;
END_VAR
END_METHOD

(* ---- L_MC4P_KINEMATIKPARAM.fb ---- *)
FUNCTION_BLOCK L_MC4P_KINEMATIKPARAM
VAR_INPUT
	ITFEXTKINPARAM : L_MC4P_IKinParamExtern;
END_VAR
END_FUNCTION_BLOCK

METHOD CALCULATEPARAMETER
END_METHOD

METHOD CHECKPARAMETER : BOOL
END_METHOD

(* ---- L_MC4P_LIMITDYNAMICSAUXAXES.fb ---- *)
FUNCTION_BLOCK L_MC4P_LIMITDYNAMICSAUXAXES EXTENDS L_MC4P_LimitDynamicsAxes
VAR_INPUT
	XENABLE : BOOL;
	ALRMAXAXESVEL : ARRAY [1..6] OF LREAL;
	ALRMAXAXESACC : ARRAY [1..6] OF LREAL;
	ALRMAXAXESJERK : ARRAY [1..6] OF LREAL;
END_VAR
VAR_OUTPUT
	XVALID : BOOL;
	XBUSY : BOOL;
	XERROR : BOOL;
	EERRORID : L_IE1P_Error := L_IE1P_Error.NoError;
END_VAR
END_FUNCTION_BLOCK

(* ---- L_MC4P_LIMITDYNAMICSAXES.fb ---- *)
FUNCTION_BLOCK L_MC4P_LIMITDYNAMICSAXES EXTENDS L_MC4P_Template_AG_KIN
VAR
	XENABLEOLD : BOOL;
	IDX : WORD;
END_VAR
END_FUNCTION_BLOCK

METHOD MAIN
VAR_INPUT
	XENABLE : BOOL;
	ALRMAXAXESVEL : ARRAY [1..6] OF LREAL;
	ALRMAXAXESACC : ARRAY [1..6] OF LREAL;
	ALRMAXAXESJERK : ARRAY [1..6] OF LREAL;
	AXESOFFSET : WORD;
END_VAR
VAR_OUTPUT
	XVALID : BOOL;
	XBUSY : BOOL;
	XERROR : BOOL;
	EERRORID : L_IE1P_Error := L_IE1P_Error.NoError;
END_VAR
VAR_IN_OUT
	AXESGROUP : AXES_GROUP_KIN;
END_VAR
END_METHOD

(* ---- L_MC4P_LIMITDYNAMICSMAINAXES.fb ---- *)
FUNCTION_BLOCK L_MC4P_LIMITDYNAMICSMAINAXES EXTENDS L_MC4P_LimitDynamicsAxes
VAR_INPUT
	XENABLE : BOOL;
	ALRMAXAXESVEL : ARRAY [1..6] OF LREAL;
	ALRMAXAXESACC : ARRAY [1..6] OF LREAL;
	ALRMAXAXESJERK : ARRAY [1..6] OF LREAL;
END_VAR
VAR_OUTPUT
	XVALID : BOOL;
	XBUSY : BOOL;
	XERROR : BOOL;
	EERRORID : L_IE1P_Error := L_IE1P_Error.NoError;
END_VAR
END_FUNCTION_BLOCK

(* ---- L_MC4P_LIMITDYNAMICSREALAXES.fb ---- *)
FUNCTION_BLOCK L_MC4P_LIMITDYNAMICSREALAXES EXTENDS L_MC4P_LimitDynamicsAxes
VAR_INPUT
	XENABLE : BOOL;
	ALRMAXAXESVEL : ARRAY [1..6] OF LREAL;
	ALRMAXAXESACC : ARRAY [1..6] OF LREAL;
	ALRMAXAXESJERK : ARRAY [1..6] OF LREAL;
END_VAR
VAR_OUTPUT
	XVALID : BOOL;
	XBUSY : BOOL;
	XERROR : BOOL;
	EERRORID : L_IE1P_Error := L_IE1P_Error.NoError;
END_VAR
END_FUNCTION_BLOCK

(* ---- L_MC4P_LISTELMINFO.fb ---- *)
FUNCTION_BLOCK L_MC4P_LISTELMINFO
VAR_INPUT
	XENABLE : BOOL;
	UDIELMIDX : UDINT := 1;
END_VAR
VAR_OUTPUT
	XBUSY : BOOL;
	XERROR : BOOL;
	EERRORID : L_IE1P_Error;
	XVALIDELM : BOOL;
	LRVMAX : LREAL;
	LRAMAX : LREAL;
	LRDMAX : LREAL;
	LRJMAX : LREAL;
	ORIGIN_X0 : ARRAY [1..6] OF LREAL;
	ORIGIN_X1 : ARRAY [1..6] OF LREAL;
	ORIGIN_X0_PTP : ARRAY [1..6] OF LREAL;
	ORIGIN_X1_PTP : ARRAY [1..6] OF LREAL;
	X0 : ARRAY [1..6] OF LREAL;
	X1 : ARRAY [1..6] OF LREAL;
	X0_PTP : ARRAY [1..6] OF LREAL;
	X1_PTP : ARRAY [1..6] OF LREAL;
	PPROFILEDATAXYZ : POINTER TO L_MC1P_ProfileData;
	DWMASK : L_MC4P_ModulMask;
END_VAR
VAR_IN_OUT
	AXESGROUP : AXES_GROUP_KIN;
END_VAR
VAR
	_MODEL : L_UBUP_BehaviourModel_LConC;
END_VAR
END_FUNCTION_BLOCK

METHOD CYCLICACTION
VAR_INPUT
	ITFTIMINGCONTROLLER : L_UBUP_ITimingController;
END_VAR
VAR_OUTPUT
	XCOMPLETE : BOOL;
	XABORT : BOOL;
	IERRORID : INT;
END_VAR
END_METHOD

METHOD FINALIZEACTION
VAR_INPUT
	XABORTPROPOSED : BOOL;
	IERRORIDPROPOSED : INT;
END_VAR
VAR_OUTPUT
	XCOMPLETE : BOOL;
	XABORT : BOOL;
	IERRORID : INT;
END_VAR
END_METHOD

METHOD RESETACTION
VAR_OUTPUT
	XCOMPLETE : BOOL;
END_VAR
END_METHOD

METHOD STARTACTION
VAR_OUTPUT
	XCOMPLETE : BOOL;
	IERRORID : INT;
END_VAR
END_METHOD

(* ---- L_MC4P_MFUNCTIONFROMPATHREF.fb ---- *)
FUNCTION_BLOCK L_MC4P_MFUNCTIONFROMPATHREF
VAR_INPUT
	PATHREF : MC_PATH_REF;
	XENABLE : BOOL;
	WMFUNCTION : WORD;
END_VAR
VAR_OUTPUT
	XBUSY : BOOL;
	XACTIVE : BOOL;
	XWAITINGFORMACKNOWLEDGE : BOOL;
	XERROR : BOOL;
	EERRORID : L_IE1P_Error;
	SCPARAMS : L_MC4P_MParams;
END_VAR
VAR
	REQUESTSINFO : DWORD;
	REQUESTSINFO_OLD : DWORD;
	DWRTRIG : DWORD;
	DWFTRIG : DWORD;
	XPATHREFVALID : BOOL;
	XWPATHREFID : __XWORD;
	DWPATHREFSTATUS : DWORD;
	XPATHREFERROR : BOOL;
	PELEMENT : POINTER TO L_MC4P_Parameter_MCMove;
	XIPOACTIVE : BOOL;
	XIPODONE : BOOL;
	XPARAMDIALOG : BOOL := FALSE;
	IVISUMPARAMI0 : INT := 1;
	PALRPARAMSACCESS : POINTER TO ARRAY [1..26] OF LREAL;
	ALRPARAMNAME : ARRAY [1..26] OF WSTRING := ["PA", "PB", "PC", "PD", "PE", "PF", "PG", "PH", "PI", "PJ", "PK", "PL", "PM", "PN", "PO", "PP", "PQ", "PR", "PS", "PT", "PU", "PV", "PW", "PX", "PY", "PZ"];
END_VAR
END_FUNCTION_BLOCK

METHOD CALL_ALLOCPOINTADR
END_METHOD

METHOD CALL_ERRORHANDLER
VAR_IN_OUT
	PATHREF : MC_PATH_REF;
END_VAR
END_METHOD

METHOD CALL_OUTPUT
END_METHOD

METHOD CALL_PATHREFINFO
END_METHOD

METHOD CALL_REQUESTS_EXT
END_METHOD

METHOD CALL_RESETOUTPUT
END_METHOD

METHOD CALL_STATEMACHINE
VAR_IN_OUT
	PATHREF : MC_PATH_REF;
END_VAR
END_METHOD

METHOD FB_INIT : BOOL
VAR_INPUT
	BINITRETAINS : BOOL;
	BINCOPYCODE : BOOL;
END_VAR
END_METHOD

(* ---- L_MC4P_MOVECIRCULARABSOLUTE_INTERNAL.fb ---- *)
FUNCTION_BLOCK L_MC4P_MOVECIRCULARABSOLUTE_INTERNAL EXTENDS L_MC4P_MoveContPath
VAR_INPUT
	EXECUTE : BOOL;
	CIRCMODE : L_MC4P_CircMode;
	AUXPOINT : ARRAY [1..12] OF LREAL;
	ENDPOINT : ARRAY [1..12] OF LREAL;
	PATHCHOICE : MC_CIRC_PATHCHOICE;
	VELOCITY : LREAL;
	ACCELERATION : LREAL;
	DECELERATION : LREAL;
	JERK : LREAL;
	COORDSYSTEM : L_MC4P_CoordSystem;
	BUFFERMODE : MC_BUFFER_MODE;
	TRANSITIONMODE : MC_TRANSITION_MODE;
	TRANSITIONPARAMETER : ARRAY [1..12] OF LREAL := [12(0)];
	AEAUXMODE : ARRAY [1..6] OF L_MC4P_AuxMode;
	ORIENTATIONMODE : L_MC4P_Orientation_Mode := L_MC4P_Orientation_Mode.ShortestSpacialWay;
	DIRECTION : ARRAY [4..6] OF MC_DIRECTION := [3(MC_DIRECTION.mcShortestWay)];
END_VAR
VAR_OUTPUT
	DONE : BOOL;
	BUSY : BOOL;
	ACTIVE : BOOL;
	COMMANDABORTED : BOOL;
	ERROR : BOOL;
	ERRORID : L_IE1P_Error;
END_VAR
VAR
	CLASSID : DINT;
END_VAR
END_FUNCTION_BLOCK

METHOD HOMINGREQUIRED : BOOL
END_METHOD

METHOD MAIN
VAR_IN_OUT
	AXESGROUP : AXES_GROUP_KIN;
	FBBASE : L_MC4P_Template_AG_KIN;
END_VAR
END_METHOD

METHOD PARAMETERFREEZE
VAR_IN_OUT
	AXESGROUP : AXES_GROUP_KIN;
	FBBASE : L_MC4P_Template_AG_KIN;
	COORDSYSTEM : L_MC4P_CoordSystem;
	BUFFERMODE : MC_BUFFER_MODE;
	TRANSITIONMODE : MC_TRANSITION_MODE;
	TRANSITIONPARAMETER : ARRAY [1..12] OF LREAL;
END_VAR
END_METHOD

METHOD SETERRORINPUTLIMITATIONVIOLATION
VAR_IN_OUT
	FBBASE : L_MC4P_Template_AG_KIN;
END_VAR
END_METHOD

METHOD SETPATHELEMENT
VAR_IN_OUT
	AXESGROUP : AXES_GROUP_KIN;
	FBBASE : L_MC4P_Template_AG_KIN;
	ALRSTARTPOS : ARRAY [1..12] OF LREAL;
	ALRSUPERPOSPOSATSTART : ARRAY [1..3] OF LREAL;
END_VAR
END_METHOD

(* ---- L_MC4P_MOVECIRCULARRELATIVE_INTERNAL.fb ---- *)
FUNCTION_BLOCK L_MC4P_MOVECIRCULARRELATIVE_INTERNAL EXTENDS L_MC4P_MoveContPath
VAR_INPUT
	EXECUTE : BOOL;
	CIRCMODE : L_MC4P_CircMode;
	AUXPOINT : ARRAY [1..12] OF LREAL;
	ENDPOINT : ARRAY [1..12] OF LREAL;
	PATHCHOICE : MC_CIRC_PATHCHOICE;
	VELOCITY : LREAL;
	ACCELERATION : LREAL;
	DECELERATION : LREAL;
	JERK : LREAL;
	COORDSYSTEM : L_MC4P_CoordSystem;
	BUFFERMODE : MC_BUFFER_MODE;
	TRANSITIONMODE : MC_TRANSITION_MODE;
	TRANSITIONPARAMETER : ARRAY [1..12] OF LREAL := [12(0)];
	AEAUXMODE : ARRAY [1..6] OF L_MC4P_AuxMode;
	ORIENTATIONMODE : L_MC4P_Orientation_Mode := L_MC4P_Orientation_Mode.ShortestSpacialWay;
	DIRECTION : ARRAY [4..6] OF MC_DIRECTION := [3(MC_DIRECTION.mcShortestWay)];
END_VAR
VAR_OUTPUT
	DONE : BOOL;
	BUSY : BOOL;
	ACTIVE : BOOL;
	COMMANDABORTED : BOOL;
	ERROR : BOOL;
	ERRORID : L_IE1P_Error;
END_VAR
VAR
	CLASSID : DINT;
END_VAR
END_FUNCTION_BLOCK

METHOD HOMINGREQUIRED : BOOL
END_METHOD

METHOD MAIN
VAR_IN_OUT
	AXESGROUP : AXES_GROUP_KIN;
	FBBASE : L_MC4P_Template_AG_KIN;
END_VAR
END_METHOD

METHOD PARAMETERFREEZE
VAR_IN_OUT
	AXESGROUP : AXES_GROUP_KIN;
	FBBASE : L_MC4P_Template_AG_KIN;
	COORDSYSTEM : L_MC4P_CoordSystem;
	BUFFERMODE : MC_BUFFER_MODE;
	TRANSITIONMODE : MC_TRANSITION_MODE;
	TRANSITIONPARAMETER : ARRAY [1..12] OF LREAL;
END_VAR
END_METHOD

METHOD SETERRORINPUTLIMITATIONVIOLATION
VAR_IN_OUT
	FBBASE : L_MC4P_Template_AG_KIN;
END_VAR
END_METHOD

METHOD SETPATHELEMENT
VAR_IN_OUT
	AXESGROUP : AXES_GROUP_KIN;
	FBBASE : L_MC4P_Template_AG_KIN;
	ALRSTARTPOS : ARRAY [1..12] OF LREAL;
	ALRSUPERPOSPOSATSTART : ARRAY [1..3] OF LREAL;
END_VAR
END_METHOD

(* ---- L_MC4P_MOVECONTPATH.fb ---- *)
FUNCTION_BLOCK L_MC4P_MOVECONTPATH EXTENDS L_UBUP_PoolInstance
VAR_INPUT
	LRCONVEYORPOSEXTRAPOL : LREAL;
	XDONTCALCPROFILEMOVEPATH : BOOL;
	ITFPATHELMDELETE : L_MC4P_IPathElmDelete;
	ITFTOOLINFO : L_MC4P_IToolInfo;
	ESRCOFCMD : L_MC4P_SourceOfMotionCommand := L_MC4P_SourceOfMotionCommand.ContPathPrepare;
END_VAR
VAR
	CALCSTOPPROFILES : L_MC4P_CalcStopProfiles;
	XMOVEREL : BOOL;
	XDONTCHECKTARGETPOSSWLIMITS : BOOL;
	XDONE_INTERN : BOOL;
	XBUSY_INTERN : BOOL;
	XACTIVE_INTERN : BOOL;
	XCOMMANDABORTED_INTERN : BOOL;
	XERROR_INTERN : BOOL;
	EERRORID_INTERN : L_IE1P_Error;
	INPUT_PARAMETER : L_MC4P_Parameter_MCMove;
	COORDTRAFOPCSFORTMPUSE : L_MC4P_CoordTrafo;
	SCPATHELEMENT : L_MC4P_PathElement;
	DIFUNID : DINT := -1;
	EXECUTEOLD : BOOL;
	WSTEP : L_MC4P_MoveContStates := L_MC4P_MoveContStates.Initial;
	WSTEPOLD : L_MC4P_MoveContStates := L_MC4P_MoveContStates.Initial;
	ALRSTARTPOS : ARRAY [1..12] OF LREAL;
	ALRPOSITIONATEXECUTE : ARRAY [1..18] OF LREAL;
	BSTATEMACHINE : BOOL;
	IPO_DONE : BOOL;
	WMASTEROFIPO : WORD;
	ERROROLD : BOOL;
	XRESETOUTPUT : BOOL := FALSE;
	SINSTANCESTR : STRING;
	ISPLINEPOINTPASSED_INTERN : INT;
	XINITABORTING : BOOL;
	PTRACKINGPARAM : POINTER TO L_MC4P_PCSTrackParam;
	PSCHANDSHAKE : POINTER TO L_MC4P_TrackingHandshake;
	XWINSTANCE : __XWORD;
	XMOVEPATHEXECUTE : BOOL;
	PSCPARMOVEPATH : POINTER TO L_MC4P_Parameter_MCMove;
	XTIMEIPOACTIVE : BOOL;
	LRCIRCANGLEEXTENDED : LREAL;
	CLASSID : DINT;
	TARGETREACHED : BOOL;
END_VAR
END_FUNCTION_BLOCK

METHOD CALCTARGETPOSITION : L_IE1P_Error
VAR_INPUT
	COORDSYSTEM : L_MC4P_CoordSystem;
	XCALCACSPOS : BOOL;
END_VAR
VAR_IN_OUT
	AXESGROUP : AXES_GROUP_KIN;
	FBBASE : L_MC4P_Template_AG_KIN;
	ALRSTARTPOS : ARRAY [1..12] OF LREAL;
	ALRPOS : ARRAY [1..12] OF LREAL;
	ALRTARGETPOS : ARRAY [1..12] OF LREAL;
	ALRTARGETPOSAUX : ARRAY [1..6] OF LREAL;
	SCTRAFOINFO : L_MC4P_TrafoInfo;
END_VAR
END_METHOD

METHOD CHECKIPOVALUES : BOOL
VAR_INPUT
	LRVELTOCHECK : LREAL;
	LRACCTOCHECK : LREAL;
	LRMAXVEL : LREAL;
	LRMAXACCDEC : LREAL;
	LRMAXJERK : LREAL;
END_VAR
VAR_IN_OUT
	AXESGROUP : AXES_GROUP_KIN;
END_VAR
END_METHOD

METHOD FB_INIT : BOOL
VAR_INPUT
	BINITRETAINS : BOOL;
	BINCOPYCODE : BOOL;
END_VAR
END_METHOD

METHOD GETPROFILETIME : LREAL
VAR_IN_OUT
	AXESGROUP : AXES_GROUP_KIN;
END_VAR
END_METHOD

METHOD GETREMAININGSEGMENTLENGTH : LREAL
VAR_IN_OUT
	AXESGROUP : AXES_GROUP_KIN;
END_VAR
END_METHOD

METHOD GETREMAININGSEGMENTTIME : BOOL
VAR_INPUT
	LRDISTANCETOTARGET : LREAL;
END_VAR
VAR_OUTPUT
	LRREMAININGTIME : LREAL;
END_VAR
VAR_IN_OUT
	AXESGROUP : AXES_GROUP_KIN;
END_VAR
END_METHOD

METHOD HOMINGREQUIRED : BOOL
END_METHOD

METHOD ISPTP : BOOL
END_METHOD

METHOD LIMITCP2AXESGROUPLIMITS : L_IE1P_Error
VAR_INPUT
	EPATHVELERRORID : L_IE1P_Error;
	EPATHACCERRORID : L_IE1P_Error;
	EPATHDECERRORID : L_IE1P_Error;
	EPATHJERKERRORID : L_IE1P_Error;
	EROTVELERRORID : L_IE1P_Error;
	EROTACCERRORID : L_IE1P_Error;
	EROTJERKERRORID : L_IE1P_Error;
	ETRANSPARAERRORID : L_IE1P_Error;
	ETRANSMODEERRORID : L_IE1P_Error;
END_VAR
VAR_IN_OUT
	AXESGROUP : AXES_GROUP_KIN;
	FBBASE : L_MC4P_Template_AG_KIN;
	AEAUXMODE : ARRAY [1..6] OF L_MC4P_AuxMode;
END_VAR
END_METHOD

METHOD PARAMETERFREEZE
VAR_IN_OUT
	AXESGROUP : AXES_GROUP_KIN;
	FBBASE : L_MC4P_Template_AG_KIN;
	COORDSYSTEM : L_MC4P_CoordSystem;
	BUFFERMODE : MC_BUFFER_MODE;
	TRANSITIONMODE : MC_TRANSITION_MODE;
	TRANSITIONPARAMETER : ARRAY [1..12] OF LREAL;
END_VAR
END_METHOD

METHOD SETERRORINPUTLIMITATIONVIOLATION
VAR_IN_OUT
	FBBASE : L_MC4P_Template_AG_KIN;
END_VAR
END_METHOD

METHOD SETPATHELEMENT_CARTESIAN
VAR_IN_OUT
	AXESGROUP : AXES_GROUP_KIN;
	FBBASE : L_MC4P_Template_AG_KIN;
	ALRSTARTPOS : ARRAY [1..12] OF LREAL;
	ALRSUPERPOSPOSATSTART : ARRAY [1..3] OF LREAL;
	AEAUXMODE : ARRAY [1..6] OF L_MC4P_AuxMode;
END_VAR
END_METHOD

METHOD SETIPO_DONE
VAR_INPUT
	IPO_DONE : BOOL;
END_VAR
END_METHOD

METHOD SETINSTANCESTRING
VAR_INPUT
	SINSTANCESTR_FATHER : STRING;
END_VAR
END_METHOD

METHOD SETMASTEROFIPO
VAR_INPUT
	WSETMASTEROFIPO : WORD;
END_VAR
END_METHOD

METHOD SETMOVECONTSTATE
VAR_INPUT
	WNEWSTEP : L_MC4P_MoveContStates;
END_VAR
END_METHOD

METHOD SETTIMEIPOACTIVEFLAG
VAR_INPUT
	XACTIVE : BOOL;
END_VAR
END_METHOD

METHOD GET_EERRORID : L_IE1P_Error
END_METHOD

METHOD GET_XACTIVE : BOOL
END_METHOD

METHOD GET_XBUSY : BOOL
END_METHOD

METHOD GET_XCOMMANDABORTED : BOOL
END_METHOD

METHOD GET_XDONE : BOOL
END_METHOD

METHOD GET_XINITIAL : BOOL
END_METHOD

METHOD FREE : BOOL
END_METHOD

METHOD REQUESTINTERFACE : BOOL
VAR_INPUT
	ID : DINT;
	PITFUNKNOWN : POINTER TO L_UBUP_IUnknown;
END_VAR
END_METHOD

METHOD CALCCIRCULARBORDERMODE : L_IE1P_Error
VAR_IN_OUT
	AXESGROUP : AXES_GROUP_KIN;
	FBBASE : L_MC4P_Template_AG_KIN;
END_VAR
END_METHOD

METHOD CALCCIRCULARCENTERMODE : L_IE1P_Error
VAR_INPUT
	ALRSTARTPOS : ARRAY [1..12] OF LREAL;
END_VAR
VAR_IN_OUT
	AXESGROUP : AXES_GROUP_KIN;
	FBBASE : L_MC4P_Template_AG_KIN;
END_VAR
END_METHOD

METHOD CALCCIRCULARRADIUSMODE : L_IE1P_Error
VAR_INPUT
	ALRSTARTPOS : ARRAY [1..12] OF LREAL;
END_VAR
VAR_IN_OUT
	AXESGROUP : AXES_GROUP_KIN;
	FBBASE : L_MC4P_Template_AG_KIN;
END_VAR
END_METHOD

METHOD SETPATHELEMENT_CIRCULAR
VAR_IN_OUT
	AXESGROUP : AXES_GROUP_KIN;
	FBBASE : L_MC4P_Template_AG_KIN;
	ALRSTARTPOS : ARRAY [1..12] OF LREAL;
	ALRSUPERPOSPOSATSTART : ARRAY [1..3] OF LREAL;
	AEAUXMODE : ARRAY [1..6] OF L_MC4P_AuxMode;
END_VAR
END_METHOD

METHOD SETPATHELEMENT_DIRECT
VAR_IN_OUT
	AXESGROUP : AXES_GROUP_KIN;
	FBBASE : L_MC4P_Template_AG_KIN;
	ALRSTARTPOS : ARRAY [1..12] OF LREAL;
	ALRSUPERPOSPOSATSTART : ARRAY [1..3] OF LREAL;
	AEAUXMODE : ARRAY [1..6] OF L_MC4P_AuxMode;
END_VAR
END_METHOD

METHOD CALCELLIPSE180DEG : L_IE1P_Error
VAR_INPUT
	ALRSTARTPOS : ARRAY [1..12] OF LREAL;
END_VAR
END_METHOD

METHOD CALCELLIPSE90DEG : L_IE1P_Error
VAR_INPUT
	ALRSTARTPOS : ARRAY [1..12] OF LREAL;
END_VAR
END_METHOD

METHOD CALCELLIPSECENTERMODE : L_IE1P_Error
VAR_INPUT
	ALRSTARTPOS : ARRAY [1..12] OF LREAL;
END_VAR
END_METHOD

METHOD SETPATHELEMENT_ELLIPTICAL
VAR_IN_OUT
	AXESGROUP : AXES_GROUP_KIN;
	FBBASE : L_MC4P_Template_AG_KIN;
	ALRSTARTPOS : ARRAY [1..12] OF LREAL;
	ALRSUPERPOSPOSATSTART : ARRAY [1..3] OF LREAL;
	AEAUXMODE : ARRAY [1..6] OF L_MC4P_AuxMode;
END_VAR
END_METHOD

METHOD SETPATHELEMENT_ELLIPTICALPNP
VAR_IN_OUT
	AXESGROUP : AXES_GROUP_KIN;
	FBBASE : L_MC4P_Template_AG_KIN;
	ALRSTARTPOS : ARRAY [1..12] OF LREAL;
	ALRSUPERPOSPOSATSTART : ARRAY [1..3] OF LREAL;
	AEAUXMODE : ARRAY [1..6] OF L_MC4P_AuxMode;
END_VAR
END_METHOD

METHOD SETPATHELEMENT_LINEAR
VAR_IN_OUT
	AXESGROUP : AXES_GROUP_KIN;
	FBBASE : L_MC4P_Template_AG_KIN;
	ALRSTARTPOS : ARRAY [1..12] OF LREAL;
	ALRSUPERPOSPOSATSTART : ARRAY [1..3] OF LREAL;
	AEAUXMODE : ARRAY [1..6] OF L_MC4P_AuxMode;
END_VAR
END_METHOD

METHOD MOVEMCMOVEPATH
VAR_IN_OUT
	XPAUSE : BOOL;
	AXESGROUP : AXES_GROUP_KIN;
	FBBASE : L_MC4P_Template_AG_KIN;
	SCPARMOVEPATH : L_MC4P_Parameter_MCMove;
	XDONE : BOOL;
	XBUSY : BOOL;
	XACTIVE : BOOL;
	XCOMMANDABORTED : BOOL;
	XERROR : BOOL;
	EERRORID : L_IE1P_Error;
END_VAR
END_METHOD

METHOD MOVEPATHDECODECIRCULAR
VAR_IN_OUT
	AXESGROUP : AXES_GROUP_KIN;
	FBBASE : L_MC4P_Template_AG_KIN;
	ALRSTARTPOS : ARRAY [1..12] OF LREAL;
END_VAR
END_METHOD

METHOD MOVEPATHINPUT
VAR_IN_OUT
	SCPARMOVEPATH : L_MC4P_Parameter_MCMove;
END_VAR
END_METHOD

METHOD PARAMETERFREEZE_MOVEPATH
VAR_IN_OUT
	AXESGROUP : AXES_GROUP_KIN;
	FBBASE : L_MC4P_Template_AG_KIN;
END_VAR
END_METHOD

METHOD SETPATHELEMENT
VAR_IN_OUT
	AXESGROUP : AXES_GROUP_KIN;
	FBBASE : L_MC4P_Template_AG_KIN;
	ALRSTARTPOS : ARRAY [1..12] OF LREAL;
	ALRSUPERPOSPOSATSTART : ARRAY [1..3] OF LREAL;
END_VAR
END_METHOD

METHOD CHECKPOINTS : L_IE1P_Error
VAR_IN_OUT
	ALRSTARTPOS : ARRAY [1..12] OF LREAL;
END_VAR
END_METHOD

METHOD PRECALCPOINTS : L_IE1P_Error
VAR_IN_OUT
	ALRSTARTPOS : ARRAY [1..12] OF LREAL;
	AXESGROUP : AXES_GROUP_KIN;
	FBBASE : L_MC4P_Template_AG_KIN;
END_VAR
END_METHOD

METHOD SETPATHELEMENT_SPLINE
VAR_IN_OUT
	AXESGROUP : AXES_GROUP_KIN;
	FBBASE : L_MC4P_Template_AG_KIN;
	ALRSTARTPOS : ARRAY [1..12] OF LREAL;
	ALRSUPERPOSPOSATSTART : ARRAY [1..3] OF LREAL;
	AEAUXMODE : ARRAY [1..6] OF L_MC4P_AuxMode;
END_VAR
END_METHOD

METHOD SETPATHELEMENT_SPLINEPNP
VAR_IN_OUT
	AXESGROUP : AXES_GROUP_KIN;
	FBBASE : L_MC4P_Template_AG_KIN;
	ALRSTARTPOS : ARRAY [1..12] OF LREAL;
	ALRSUPERPOSPOSATSTART : ARRAY [1..3] OF LREAL;
	AEAUXMODE : ARRAY [1..6] OF L_MC4P_AuxMode;
END_VAR
END_METHOD

METHOD SETSPLINEPOINTPASSED
VAR_INPUT
	UIPOINTPASSED : UINT;
END_VAR
END_METHOD

METHOD MOVECONTPATH
VAR_IN_OUT
	AXESGROUP : AXES_GROUP_KIN;
	FBBASE : L_MC4P_Template_AG_KIN;
	EXECUTE : BOOL;
	COORDSYSTEM : L_MC4P_CoordSystem;
	AEAUXMODE : ARRAY [1..6] OF L_MC4P_AuxMode;
	BUFFERMODE : MC_BUFFER_MODE;
	TRANSITIONMODE : MC_TRANSITION_MODE;
	TRANSITIONPARAMETER : ARRAY [1..12] OF LREAL;
END_VAR
END_METHOD

METHOD MOVECONTSTATES_ABORTING
VAR_IN_OUT
	AXESGROUP : AXES_GROUP_KIN;
	FBBASE : L_MC4P_Template_AG_KIN;
	EXECUTE : BOOL;
	COORDSYSTEM : L_MC4P_CoordSystem;
	AEAUXMODE : ARRAY [1..6] OF L_MC4P_AuxMode;
	BUFFERMODE : MC_BUFFER_MODE;
	TRANSITIONMODE : MC_TRANSITION_MODE;
	TRANSITIONPARAMETER : ARRAY [1..12] OF LREAL;
END_VAR
END_METHOD

METHOD MOVECONTSTATES_CALCPATH
VAR_IN_OUT
	AXESGROUP : AXES_GROUP_KIN;
	FBBASE : L_MC4P_Template_AG_KIN;
	EXECUTE : BOOL;
	COORDSYSTEM : L_MC4P_CoordSystem;
	AEAUXMODE : ARRAY [1..6] OF L_MC4P_AuxMode;
	BUFFERMODE : MC_BUFFER_MODE;
	TRANSITIONMODE : MC_TRANSITION_MODE;
	TRANSITIONPARAMETER : ARRAY [1..12] OF LREAL;
END_VAR
END_METHOD

METHOD MOVECONTSTATES_ERRORSTATE
VAR_IN_OUT
	AXESGROUP : AXES_GROUP_KIN;
	FBBASE : L_MC4P_Template_AG_KIN;
	EXECUTE : BOOL;
	COORDSYSTEM : L_MC4P_CoordSystem;
	AEAUXMODE : ARRAY [1..6] OF L_MC4P_AuxMode;
	BUFFERMODE : MC_BUFFER_MODE;
	TRANSITIONMODE : MC_TRANSITION_MODE;
	TRANSITIONPARAMETER : ARRAY [1..12] OF LREAL;
END_VAR
END_METHOD

METHOD MOVECONTSTATES_IPO_ACTIVE
VAR_IN_OUT
	AXESGROUP : AXES_GROUP_KIN;
	FBBASE : L_MC4P_Template_AG_KIN;
	EXECUTE : BOOL;
	COORDSYSTEM : L_MC4P_CoordSystem;
	AEAUXMODE : ARRAY [1..6] OF L_MC4P_AuxMode;
	BUFFERMODE : MC_BUFFER_MODE;
	TRANSITIONMODE : MC_TRANSITION_MODE;
	TRANSITIONPARAMETER : ARRAY [1..12] OF LREAL;
END_VAR
END_METHOD

METHOD MOVECONTSTATES_IPO_STANDBY
VAR_IN_OUT
	AXESGROUP : AXES_GROUP_KIN;
	FBBASE : L_MC4P_Template_AG_KIN;
	EXECUTE : BOOL;
	COORDSYSTEM : L_MC4P_CoordSystem;
	AEAUXMODE : ARRAY [1..6] OF L_MC4P_AuxMode;
	BUFFERMODE : MC_BUFFER_MODE;
	TRANSITIONMODE : MC_TRANSITION_MODE;
	TRANSITIONPARAMETER : ARRAY [1..12] OF LREAL;
END_VAR
END_METHOD

METHOD MOVECONTSTATES_INITIAL
VAR_IN_OUT
	AXESGROUP : AXES_GROUP_KIN;
	FBBASE : L_MC4P_Template_AG_KIN;
	EXECUTE : BOOL;
	COORDSYSTEM : L_MC4P_CoordSystem;
	AEAUXMODE : ARRAY [1..6] OF L_MC4P_AuxMode;
	BUFFERMODE : MC_BUFFER_MODE;
	TRANSITIONMODE : MC_TRANSITION_MODE;
	TRANSITIONPARAMETER : ARRAY [1..12] OF LREAL;
END_VAR
END_METHOD

METHOD MOVECONTSTATES_READPARAM_STANDBY
VAR_IN_OUT
	AXESGROUP : AXES_GROUP_KIN;
	FBBASE : L_MC4P_Template_AG_KIN;
	EXECUTE : BOOL;
	COORDSYSTEM : L_MC4P_CoordSystem;
	AEAUXMODE : ARRAY [1..6] OF L_MC4P_AuxMode;
	BUFFERMODE : MC_BUFFER_MODE;
	TRANSITIONMODE : MC_TRANSITION_MODE;
	TRANSITIONPARAMETER : ARRAY [1..12] OF LREAL;
END_VAR
END_METHOD

METHOD MOVECONTSTATES_READ_INPUTS
VAR_IN_OUT
	AXESGROUP : AXES_GROUP_KIN;
	FBBASE : L_MC4P_Template_AG_KIN;
	EXECUTE : BOOL;
	COORDSYSTEM : L_MC4P_CoordSystem;
	AEAUXMODE : ARRAY [1..6] OF L_MC4P_AuxMode;
	BUFFERMODE : MC_BUFFER_MODE;
	TRANSITIONMODE : MC_TRANSITION_MODE;
	TRANSITIONPARAMETER : ARRAY [1..12] OF LREAL;
END_VAR
END_METHOD

METHOD SETPATHELEMENT_WAITTIME
VAR_IN_OUT
	AXESGROUP : AXES_GROUP_KIN;
	FBBASE : L_MC4P_Template_AG_KIN;
	ALRSTARTPOS : ARRAY [1..12] OF LREAL;
	ALRSUPERPOSPOSATSTART : ARRAY [1..3] OF LREAL;
	LRWAITTIME : LREAL;
	EERRORID : L_IE1P_Error;
END_VAR
END_METHOD

(* ---- L_MC4P_MOVEDIRECTABSOLUTE_INTERNAL.fb ---- *)
FUNCTION_BLOCK L_MC4P_MOVEDIRECTABSOLUTE_INTERNAL EXTENDS L_MC4P_MoveContPath
VAR_INPUT
	EXECUTE : BOOL;
	POSITION : ARRAY [1..12] OF LREAL;
	COORDSYSTEM : L_MC4P_CoordSystem;
	BUFFERMODE : MC_BUFFER_MODE;
	TRANSITIONMODE : MC_TRANSITION_MODE;
	TRANSITIONPARAMETER : ARRAY [1..12] OF LREAL := [12(0)];
	AITARGETCONFIGURATION : ARRAY [1..6] OF INT;
	DIRECTION : ARRAY [1..6] OF MC_DIRECTION := [6(MC_DIRECTION.mcShortestWay)];
END_VAR
VAR_OUTPUT
	DONE : BOOL;
	BUSY : BOOL;
	ACTIVE : BOOL;
	COMMANDABORTED : BOOL;
	ERROR : BOOL;
	ERRORID : L_IE1P_Error;
END_VAR
VAR
	AEAUXMODE : ARRAY [1..6] OF L_MC4P_AuxMode := [6(L_MC4P_AuxMode.Inactive)];
	CLASSID : DINT;
END_VAR
END_FUNCTION_BLOCK

METHOD HOMINGREQUIRED : BOOL
END_METHOD

METHOD ISPTP : BOOL
END_METHOD

METHOD MAIN
VAR_IN_OUT
	AXESGROUP : AXES_GROUP_KIN;
	FBBASE : L_MC4P_Template_AG_KIN;
END_VAR
END_METHOD

METHOD PARAMETERFREEZE
VAR_IN_OUT
	AXESGROUP : AXES_GROUP_KIN;
	FBBASE : L_MC4P_Template_AG_KIN;
	COORDSYSTEM : L_MC4P_CoordSystem;
	BUFFERMODE : MC_BUFFER_MODE;
	TRANSITIONMODE : MC_TRANSITION_MODE;
	TRANSITIONPARAMETER : ARRAY [1..12] OF LREAL;
END_VAR
END_METHOD

METHOD SETERRORINPUTLIMITATIONVIOLATION
VAR_IN_OUT
	FBBASE : L_MC4P_Template_AG_KIN;
END_VAR
END_METHOD

METHOD SETPATHELEMENT
VAR_IN_OUT
	AXESGROUP : AXES_GROUP_KIN;
	FBBASE : L_MC4P_Template_AG_KIN;
	ALRSTARTPOS : ARRAY [1..12] OF LREAL;
	ALRSUPERPOSPOSATSTART : ARRAY [1..3] OF LREAL;
END_VAR
END_METHOD

(* ---- L_MC4P_MOVEDIRECTRELATIVE_INTERNAL.fb ---- *)
FUNCTION_BLOCK L_MC4P_MOVEDIRECTRELATIVE_INTERNAL EXTENDS L_MC4P_MoveContPath
VAR_INPUT
	EXECUTE : BOOL;
	DISTANCE : ARRAY [1..12] OF LREAL;
	COORDSYSTEM : L_MC4P_CoordSystem;
	BUFFERMODE : MC_BUFFER_MODE;
	TRANSITIONMODE : MC_TRANSITION_MODE;
	TRANSITIONPARAMETER : ARRAY [1..12] OF LREAL := [12(0)];
	AITARGETCONFIGURATION : ARRAY [1..6] OF INT;
	DIRECTION : ARRAY [1..6] OF MC_DIRECTION := [6(MC_DIRECTION.mcShortestWay)];
END_VAR
VAR_OUTPUT
	DONE : BOOL;
	BUSY : BOOL;
	ACTIVE : BOOL;
	COMMANDABORTED : BOOL;
	ERROR : BOOL;
	ERRORID : L_IE1P_Error;
END_VAR
VAR
	AEAUXMODE : ARRAY [1..6] OF L_MC4P_AuxMode := [6(L_MC4P_AuxMode.Inactive)];
	CLASSID : DINT;
END_VAR
END_FUNCTION_BLOCK

METHOD HOMINGREQUIRED : BOOL
END_METHOD

METHOD ISPTP : BOOL
END_METHOD

METHOD MAIN
VAR_IN_OUT
	AXESGROUP : AXES_GROUP_KIN;
	FBBASE : L_MC4P_Template_AG_KIN;
END_VAR
END_METHOD

METHOD PARAMETERFREEZE
VAR_IN_OUT
	AXESGROUP : AXES_GROUP_KIN;
	FBBASE : L_MC4P_Template_AG_KIN;
	COORDSYSTEM : L_MC4P_CoordSystem;
	BUFFERMODE : MC_BUFFER_MODE;
	TRANSITIONMODE : MC_TRANSITION_MODE;
	TRANSITIONPARAMETER : ARRAY [1..12] OF LREAL;
END_VAR
END_METHOD

METHOD SETERRORINPUTLIMITATIONVIOLATION
VAR_IN_OUT
	FBBASE : L_MC4P_Template_AG_KIN;
END_VAR
END_METHOD

METHOD SETPATHELEMENT
VAR_IN_OUT
	AXESGROUP : AXES_GROUP_KIN;
	FBBASE : L_MC4P_Template_AG_KIN;
	ALRSTARTPOS : ARRAY [1..12] OF LREAL;
	ALRSUPERPOSPOSATSTART : ARRAY [1..3] OF LREAL;
END_VAR
END_METHOD

(* ---- L_MC4P_MOVEELLIPTICALABSOLUTE.fb ---- *)
FUNCTION_BLOCK L_MC4P_MOVEELLIPTICALABSOLUTE EXTENDS L_MC4P_Template_MoveLicence
VAR_INPUT
	XEXECUTE : BOOL;
	ALRAUXPOINT : ARRAY [1..12] OF LREAL;
	ALRENDPOINT : ARRAY [1..12] OF LREAL;
	LRSEMIMAJORAXIS : LREAL;
	LRSEMIMINORAXIS : LREAL;
	EPATHCHOICE : MC_CIRC_PATHCHOICE;
	LRVELOCITY : LREAL;
	LRACCELERATION : LREAL;
	LRDECELERATION : LREAL;
	LRJERK : LREAL;
	ECOORDSYSTEM : L_MC4P_CoordSystem;
	EBUFFERMODE : MC_BUFFER_MODE;
	ETRANSITIONMODE : MC_TRANSITION_MODE;
	ALRTRANSITIONPARAMETER : ARRAY [1..12] OF LREAL := [12(0)];
	AEAUXMODE : ARRAY [1..6] OF L_MC4P_AuxMode;
	EORIENTATIONMODE : L_MC4P_Orientation_Mode := L_MC4P_Orientation_Mode.ShortestSpacialWay;
	AEDIRECTION : ARRAY [4..6] OF MC_DIRECTION := [3(MC_DIRECTION.mcShortestWay)];
END_VAR
VAR_OUTPUT
	XDONE : BOOL;
	XBUSY : BOOL;
	XACTIVE : BOOL;
	XCOMMANDABORTED : BOOL;
	XERROR : BOOL;
	EERRORID : L_IE1P_Error;
END_VAR
VAR
	MOVEELLIPTICAL : L_MC4P_MoveEllipticalAbsolute_Internal;
	PMOVE : POINTER TO L_MC4P_MoveContPath;
	SETELLIPTICALTARGETTOLERANCE : LREAL;
END_VAR
END_FUNCTION_BLOCK

(* ---- L_MC4P_MOVEELLIPTICALABSOLUTE_INTERNAL.fb ---- *)
FUNCTION_BLOCK L_MC4P_MOVEELLIPTICALABSOLUTE_INTERNAL EXTENDS L_MC4P_MoveContPath
VAR_INPUT
	XEXECUTE : BOOL;
	ALRAUXPOINT : ARRAY [1..12] OF LREAL;
	ALRENDPOINT : ARRAY [1..12] OF LREAL;
	LRSEMIMAJORAXIS : LREAL;
	LRSEMIMINORAXIS : LREAL;
	EPATHCHOICE : MC_CIRC_PATHCHOICE;
	LRVELOCITY : LREAL;
	LRACCELERATION : LREAL;
	LRDECELERATION : LREAL;
	LRJERK : LREAL;
	ECOORDSYSTEM : L_MC4P_CoordSystem;
	EBUFFERMODE : MC_BUFFER_MODE;
	ETRANSITIONMODE : MC_TRANSITION_MODE;
	ALRTRANSITIONPARAMETER : ARRAY [1..12] OF LREAL := [12(0)];
	AEAUXMODE : ARRAY [1..6] OF L_MC4P_AuxMode;
	EORIENTATIONMODE : L_MC4P_Orientation_Mode := L_MC4P_Orientation_Mode.ShortestSpacialWay;
	AEDIRECTION : ARRAY [4..6] OF MC_DIRECTION := [3(MC_DIRECTION.mcShortestWay)];
END_VAR
VAR_OUTPUT
	XDONE : BOOL;
	XBUSY : BOOL;
	XACTIVE : BOOL;
	XCOMMANDABORTED : BOOL;
	XERROR : BOOL;
	EERRORID : L_IE1P_Error;
END_VAR
VAR
	ECIRCMODE : L_MC4P_CircMode := L_MC4P_CircMode.CENTER;
	CLASSID : DINT;
END_VAR
END_FUNCTION_BLOCK

METHOD HOMINGREQUIRED : BOOL
END_METHOD

METHOD MAIN
VAR_IN_OUT
	AXESGROUP : AXES_GROUP_KIN;
	FBBASE : L_MC4P_Template_AG_KIN;
END_VAR
END_METHOD

METHOD PARAMETERFREEZE
VAR_IN_OUT
	AXESGROUP : AXES_GROUP_KIN;
	FBBASE : L_MC4P_Template_AG_KIN;
	COORDSYSTEM : L_MC4P_CoordSystem;
	BUFFERMODE : MC_BUFFER_MODE;
	TRANSITIONMODE : MC_TRANSITION_MODE;
	TRANSITIONPARAMETER : ARRAY [1..12] OF LREAL;
END_VAR
END_METHOD

METHOD SETERRORINPUTLIMITATIONVIOLATION
VAR_IN_OUT
	FBBASE : L_MC4P_Template_AG_KIN;
END_VAR
END_METHOD

METHOD SETPATHELEMENT
VAR_IN_OUT
	AXESGROUP : AXES_GROUP_KIN;
	FBBASE : L_MC4P_Template_AG_KIN;
	ALRSTARTPOS : ARRAY [1..12] OF LREAL;
	ALRSUPERPOSPOSATSTART : ARRAY [1..3] OF LREAL;
END_VAR
END_METHOD

METHOD FB_INIT : BOOL
VAR_INPUT
	BINITRETAINS : BOOL;
	BINCOPYCODE : BOOL;
END_VAR
END_METHOD

(* ---- L_MC4P_MOVEELLIPTICALABSOLUTEPNP.fb ---- *)
FUNCTION_BLOCK L_MC4P_MOVEELLIPTICALABSOLUTEPNP EXTENDS L_MC4P_Template_MoveLicence
VAR_INPUT
	XEXECUTE : BOOL;
	ALRENDPOINT : ARRAY [1..12] OF LREAL;
	ALRDIRECTION : ARRAY [1..3] OF LREAL;
	LRSEMIAXIS : LREAL;
	EELLIPTICALPNPMODE : L_MC4P_EllipticalPnPMode := L_MC4P_EllipticalPnPMode.Elliptical_180;
	LRVELOCITY : LREAL;
	LRACCELERATION : LREAL;
	LRDECELERATION : LREAL;
	LRJERK : LREAL;
	ECOORDSYSTEM : L_MC4P_CoordSystem;
	EBUFFERMODE : MC_BUFFER_MODE;
	ETRANSITIONMODE : MC_TRANSITION_MODE;
	ALRTRANSITIONPARAMETER : ARRAY [1..12] OF LREAL := [12(0)];
	AEAUXMODE : ARRAY [1..6] OF L_MC4P_AuxMode;
	EORIENTATIONMODE : L_MC4P_Orientation_Mode := L_MC4P_Orientation_Mode.ShortestSpacialWay;
	AEDIRECTION : ARRAY [4..6] OF MC_DIRECTION := [3(MC_DIRECTION.mcShortestWay)];
END_VAR
VAR_OUTPUT
	XDONE : BOOL;
	XBUSY : BOOL;
	XACTIVE : BOOL;
	XCOMMANDABORTED : BOOL;
	XERROR : BOOL;
	EERRORID : L_IE1P_Error;
END_VAR
VAR
	MOVEELLIPTICAL : L_MC4P_MoveEllipticalAbsolutePnP_Internal;
	PMOVE : POINTER TO L_MC4P_MoveContPath;
END_VAR
END_FUNCTION_BLOCK

(* ---- L_MC4P_MOVEELLIPTICALABSOLUTEPNP_INTERNAL.fb ---- *)
FUNCTION_BLOCK L_MC4P_MOVEELLIPTICALABSOLUTEPNP_INTERNAL EXTENDS L_MC4P_MoveContPath
VAR_INPUT
	XEXECUTE : BOOL;
	ALRENDPOINT : ARRAY [1..12] OF LREAL;
	ALRDIRECTION : ARRAY [1..3] OF LREAL;
	LRSEMIAXIS : LREAL;
	EELLIPTICALPNPMODE : L_MC4P_EllipticalPnPMode := L_MC4P_EllipticalPnPMode.Elliptical_180;
	LRVELOCITY : LREAL;
	LRACCELERATION : LREAL;
	LRDECELERATION : LREAL;
	LRJERK : LREAL;
	ECOORDSYSTEM : L_MC4P_CoordSystem;
	EBUFFERMODE : MC_BUFFER_MODE;
	ETRANSITIONMODE : MC_TRANSITION_MODE;
	ALRTRANSITIONPARAMETER : ARRAY [1..12] OF LREAL := [12(0)];
	AEAUXMODE : ARRAY [1..6] OF L_MC4P_AuxMode;
	EORIENTATIONMODE : L_MC4P_Orientation_Mode := L_MC4P_Orientation_Mode.ShortestSpacialWay;
	AEDIRECTION : ARRAY [4..6] OF MC_DIRECTION := [3(MC_DIRECTION.mcShortestWay)];
END_VAR
VAR_OUTPUT
	XDONE : BOOL;
	XBUSY : BOOL;
	XACTIVE : BOOL;
	XCOMMANDABORTED : BOOL;
	XERROR : BOOL;
	EERRORID : L_IE1P_Error;
END_VAR
VAR
	ECIRCMODE : L_MC4P_CircMode := L_MC4P_CircMode.CENTER;
	EPATHCHOICE : MC_CIRC_PATHCHOICE := MC_CIRC_PATHCHOICE.CLOCKWISE;
	CLASSID : DINT;
END_VAR
END_FUNCTION_BLOCK

METHOD HOMINGREQUIRED : BOOL
END_METHOD

METHOD MAIN
VAR_IN_OUT
	AXESGROUP : AXES_GROUP_KIN;
	FBBASE : L_MC4P_Template_AG_KIN;
END_VAR
END_METHOD

METHOD PARAMETERFREEZE
VAR_IN_OUT
	AXESGROUP : AXES_GROUP_KIN;
	FBBASE : L_MC4P_Template_AG_KIN;
	COORDSYSTEM : L_MC4P_CoordSystem;
	BUFFERMODE : MC_BUFFER_MODE;
	TRANSITIONMODE : MC_TRANSITION_MODE;
	TRANSITIONPARAMETER : ARRAY [1..12] OF LREAL;
END_VAR
END_METHOD

METHOD SETERRORINPUTLIMITATIONVIOLATION
VAR_IN_OUT
	FBBASE : L_MC4P_Template_AG_KIN;
END_VAR
END_METHOD

METHOD SETPATHELEMENT
VAR_IN_OUT
	AXESGROUP : AXES_GROUP_KIN;
	FBBASE : L_MC4P_Template_AG_KIN;
	ALRSTARTPOS : ARRAY [1..12] OF LREAL;
	ALRSUPERPOSPOSATSTART : ARRAY [1..3] OF LREAL;
END_VAR
END_METHOD

METHOD FB_INIT : BOOL
VAR_INPUT
	BINITRETAINS : BOOL;
	BINCOPYCODE : BOOL;
END_VAR
END_METHOD

(* ---- L_MC4P_MOVEELLIPTICALRELATIVE.fb ---- *)
FUNCTION_BLOCK L_MC4P_MOVEELLIPTICALRELATIVE EXTENDS L_MC4P_Template_MoveLicence
VAR_INPUT
	XEXECUTE : BOOL;
	ALRAUXPOINT : ARRAY [1..12] OF LREAL;
	ALRENDPOINT : ARRAY [1..12] OF LREAL;
	LRSEMIMAJORAXIS : LREAL;
	LRSEMIMINORAXIS : LREAL;
	EPATHCHOICE : MC_CIRC_PATHCHOICE;
	LRVELOCITY : LREAL;
	LRACCELERATION : LREAL;
	LRDECELERATION : LREAL;
	LRJERK : LREAL;
	ECOORDSYSTEM : L_MC4P_CoordSystem;
	EBUFFERMODE : MC_BUFFER_MODE;
	ETRANSITIONMODE : MC_TRANSITION_MODE;
	ALRTRANSITIONPARAMETER : ARRAY [1..12] OF LREAL := [12(0)];
	AEAUXMODE : ARRAY [1..6] OF L_MC4P_AuxMode;
	EORIENTATIONMODE : L_MC4P_Orientation_Mode := L_MC4P_Orientation_Mode.ShortestSpacialWay;
	AEDIRECTION : ARRAY [4..6] OF MC_DIRECTION := [3(MC_DIRECTION.mcShortestWay)];
END_VAR
VAR_OUTPUT
	XDONE : BOOL;
	XBUSY : BOOL;
	XACTIVE : BOOL;
	XCOMMANDABORTED : BOOL;
	XERROR : BOOL;
	EERRORID : L_IE1P_Error;
END_VAR
VAR
	MOVEELLIPTICAL : L_MC4P_MoveEllipticalRelative_Internal;
	PMOVE : POINTER TO L_MC4P_MoveContPath;
	SETELLIPTICALTARGETTOLERANCE : LREAL;
END_VAR
END_FUNCTION_BLOCK

(* ---- L_MC4P_MOVEELLIPTICALRELATIVE_INTERNAL.fb ---- *)
FUNCTION_BLOCK L_MC4P_MOVEELLIPTICALRELATIVE_INTERNAL EXTENDS L_MC4P_MoveContPath
VAR_INPUT
	XEXECUTE : BOOL;
	ALRAUXPOINT : ARRAY [1..12] OF LREAL;
	ALRENDPOINT : ARRAY [1..12] OF LREAL;
	LRSEMIMAJORAXIS : LREAL;
	LRSEMIMINORAXIS : LREAL;
	EPATHCHOICE : MC_CIRC_PATHCHOICE;
	LRVELOCITY : LREAL;
	LRACCELERATION : LREAL;
	LRDECELERATION : LREAL;
	LRJERK : LREAL;
	ECOORDSYSTEM : L_MC4P_CoordSystem;
	EBUFFERMODE : MC_BUFFER_MODE;
	ETRANSITIONMODE : MC_TRANSITION_MODE;
	ALRTRANSITIONPARAMETER : ARRAY [1..12] OF LREAL := [12(0)];
	AEAUXMODE : ARRAY [1..6] OF L_MC4P_AuxMode;
	EORIENTATIONMODE : L_MC4P_Orientation_Mode := L_MC4P_Orientation_Mode.ShortestSpacialWay;
	AEDIRECTION : ARRAY [4..6] OF MC_DIRECTION := [3(MC_DIRECTION.mcShortestWay)];
END_VAR
VAR_OUTPUT
	XDONE : BOOL;
	XBUSY : BOOL;
	XACTIVE : BOOL;
	XCOMMANDABORTED : BOOL;
	XERROR : BOOL;
	EERRORID : L_IE1P_Error;
END_VAR
VAR
	ECIRCMODE : L_MC4P_CircMode := L_MC4P_CircMode.CENTER;
	CLASSID : DINT;
END_VAR
END_FUNCTION_BLOCK

METHOD HOMINGREQUIRED : BOOL
END_METHOD

METHOD MAIN
VAR_IN_OUT
	AXESGROUP : AXES_GROUP_KIN;
	FBBASE : L_MC4P_Template_AG_KIN;
END_VAR
END_METHOD

METHOD PARAMETERFREEZE
VAR_IN_OUT
	AXESGROUP : AXES_GROUP_KIN;
	FBBASE : L_MC4P_Template_AG_KIN;
	COORDSYSTEM : L_MC4P_CoordSystem;
	BUFFERMODE : MC_BUFFER_MODE;
	TRANSITIONMODE : MC_TRANSITION_MODE;
	TRANSITIONPARAMETER : ARRAY [1..12] OF LREAL;
END_VAR
END_METHOD

METHOD SETERRORINPUTLIMITATIONVIOLATION
VAR_IN_OUT
	FBBASE : L_MC4P_Template_AG_KIN;
END_VAR
END_METHOD

METHOD SETPATHELEMENT
VAR_IN_OUT
	AXESGROUP : AXES_GROUP_KIN;
	FBBASE : L_MC4P_Template_AG_KIN;
	ALRSTARTPOS : ARRAY [1..12] OF LREAL;
	ALRSUPERPOSPOSATSTART : ARRAY [1..3] OF LREAL;
END_VAR
END_METHOD

METHOD FB_INIT : BOOL
VAR_INPUT
	BINITRETAINS : BOOL;
	BINCOPYCODE : BOOL;
END_VAR
END_METHOD

(* ---- L_MC4P_MOVEFBDIAGNOSTIC.fb ---- *)
FUNCTION_BLOCK L_MC4P_MOVEFBDIAGNOSTIC
VAR_INPUT
	XEXECUTEWRITETEXTFILE : BOOL;
	XENABLE : BOOL;
END_VAR
VAR_OUTPUT
	XWRITEFILEDONE : BOOL;
	XWRITEFILEBUSY : BOOL;
	XWRITEFILEERROR : BOOL;
	XBUSY : BOOL;
END_VAR
VAR
	ASCPARAMS : ARRAY [0..wDepth] OF L_MC4P_Parameter_MCMove;
	ADWTIMESTAMP : ARRAY [0..wDepth] OF DWORD;
	ASINSTANCESTR : ARRAY [0..wDepth] OF STRING;
	WCURRENTPOS : WORD := 0;
	SCPARAMDUMMY : L_MC4P_Parameter_MCMove;
	XTESTINMOTIONTASK : BOOL := FALSE;
	XFREETASKBUSY_INT : BOOL;
	XFREETASKDONE_INT : BOOL;
	XFREETASKERROR_INT : BOOL;
	EFREETASKEERRORID_INT : L_IE1P_Error;
	XEXECUTEWRITETEXTFILE_OLD : BOOL;
	SEXCELFILENAME : STRING(255);
	RES : SYSFILE.RTS_IEC_ResULT;
	HFILE : SYSFILE.RTS_IEC_HANDLE;
	XWFSIZE : __XWORD;
	XWRESULTWRITESTRING : __XWORD;
	ASHEADLINEPARAMS : ARRAY [1..iMaxHeadLine] OF STRING := ['TimeStamp', 'sInstanceStr', 'SegmentType', 'xMoveRel', 'Position', 'Distance', 'CircMode', 'AuxPoint', 'PathChoice', 'lrSemiMajorAxis', 'lrSemiMinorAxis', 'ascIntermediatePointSpline', 'Velocity', 'Acceleration', 'Deceleration', 'Jerk', 'alrVelocityPTP', 'alrAccelerationPTP', 'alrDecelerationPTP', 'alrJerkPTP', 'alrVelocityAux', 'alrAccelerationAux', 'alrDecelerationAux', 'alrJerkAux', 'CoordSystem', 'CoordRef', 'BufferMode', 'TransitionMode', 'TransitionParameter', 'aeAuxMode', 'alrAxisLimitVel', 'alrAxisLimitAcc', 'alrAxisLimitJerk', 'aiTargetConfiguration', 'eOrientationMode', 'aeDirection'];
	STABULATOR : STRING(2) := '$T';
	SLINEFEED : STRING(2) := '$N';
	SZEILE : STRING(255);
	WSTEPWF : WORD := 0;
	XAGERROR : BOOL;
	WLOOKAHEADHORIZON : WORD;
	DWTASKCYCLE_US : DWORD;
	EACTIVEERRORID : L_IE1P_Error;
	SAXESGROUPNAME : STRING;
	VERSION : VERSION;
	WDEPTH : WORD := 50;
	IMAXHEADLINE : INT := 40;
	ACTIVEERRORID : WORD;
	AGERROR : BOOL;
	AXESGROUPNAME : STRING;
	LOOKAHEADHORIZON : WORD;
	TASKCYCLE_US : DWORD;
	VERSIONMC4P : VERSION;
	XWRITEINMOTIONTASK : BOOL;
END_VAR
END_FUNCTION_BLOCK

METHOD FREEZEMOVEFBPARAM
VAR_INPUT
	SINSTANCESTR : STRING;
	DWTIMESTAMP : DWORD;
END_VAR
VAR_IN_OUT
	INPUT_PARAMETER : L_MC4P_Parameter_MCMove;
END_VAR
END_METHOD

METHOD FREEZESTOPALLPARAM
VAR_INPUT
	SINSTANCESTR : STRING;
	DWTIMESTAMP : DWORD;
END_VAR
VAR_IN_OUT
	ASCCTRLABC : ARRAY [1..18] OF L_MC1P_CtrlABC;
END_VAR
END_METHOD

METHOD FREEZESTOPPARAM
VAR_INPUT
	SINSTANCESTR : STRING;
	DWTIMESTAMP : DWORD;
	LRINPUTDECELERATION : LREAL;
	LRINPUTJERK : LREAL;
END_VAR
END_METHOD

METHOD CALL_WRITEEXCELFILE
END_METHOD

METHOD EXECUTEFREERUNTASK
VAR_INPUT
	SDIR : STRING;
END_VAR
END_METHOD

METHOD MAIN
END_METHOD

METHOD ABORT : UDINT
END_METHOD

METHOD EXECUTE : UDINT
END_METHOD

(* ---- L_MC4P_MOVEFBPOOL.fb ---- *)
FUNCTION_BLOCK L_MC4P_MOVEFBPOOL EXTENDS L_UBUP_FBPool
VAR
	_PICKANDPLACEMEMORY : REFERENCE TO L_MC4P_PickAndPlaceMemory;
	_XMEMOWNER1 : BOOL;
	_SCFBSTORE : REFERENCE TO L_MC4P_MovePathStore;
	_XMEMOWNER2 : BOOL;
	_AFB_MOVEELLIPTICALABS : ARRAY [1..3] OF L_MC4P_MoveEllipticalAbsolute_Internal;
	_MOVELINABSCONTROLNODES : L_UBUP_DoubleLinkedListNodes;
	_MOVELINABSCONTROL : L_UBUP_DoubleLinkedListControl;
	_MOVELINRELCONTROLNODES : L_UBUP_DoubleLinkedListNodes;
	_MOVELINRELCONTROL : L_UBUP_DoubleLinkedListControl;
	_MOVEDIRABSCONTROLNODES : L_UBUP_DoubleLinkedListNodes;
	_MOVEDIRABSCONTROL : L_UBUP_DoubleLinkedListControl;
	_MOVEDIRRELCONTROLNODES : L_UBUP_DoubleLinkedListNodes;
	_MOVEDIRRELCONTROL : L_UBUP_DoubleLinkedListControl;
	_MOVEELLIPTPNPCONTROLNODES : L_UBUP_DoubleLinkedListNodes;
	_MOVEELLIPTPNPCONTROL : L_UBUP_DoubleLinkedListControl;
	_MOVEELLIPTABSCONTROLNODES : L_UBUP_DoubleLinkedListNodes;
	_MOVEELLIPTABSCONTROL : L_UBUP_DoubleLinkedListControl;
	_MOVESPLINEPNPCONTROLNODES : L_UBUP_DoubleLinkedListNodes;
	_MOVESPLINEPNPCONTROL : L_UBUP_DoubleLinkedListControl;
	_MOVECONTPATHCONTROLNODES : L_UBUP_DoubleLinkedListNodes;
	_MOVECONTPATHCONTROL : L_UBUP_DoubleLinkedListControl;
	USEGLOBAL : BOOL;
END_VAR
END_FUNCTION_BLOCK

METHOD FREEINSTANCE : BOOL
VAR_INPUT
	ITFINSTANCE : L_UBUP_IPoolInstance;
	XWHANDLE : __XWORD;
END_VAR
END_METHOD

METHOD GETCAPACITY : BOOL
VAR_INPUT
	ECLASSID : DINT;
END_VAR
VAR_OUTPUT
	DWCAPACITY : DWORD;
END_VAR
END_METHOD

METHOD QUERYINSTANCE : BOOL
VAR_INPUT
	ECLASSID : DINT;
END_VAR
VAR_IN_OUT
	ITFINSTANCE : L_UBUP_IPoolInstance;
END_VAR
END_METHOD

METHOD FB_INIT : BOOL
VAR_INPUT
	BINITRETAINS : BOOL;
	BINCOPYCODE : BOOL;
END_VAR
END_METHOD

METHOD FB_AFTERGLOBALINIT : BOOL
END_METHOD

METHOD FREERESOURCE
END_METHOD

METHOD GETFB : L_UBUP_IPoolInstance
VAR_INPUT
	ECLASSID : DINT;
	DWARRIDX : DWORD;
END_VAR
END_METHOD

METHOD GETFBCONTROL : L_UBUP_IListControl
VAR_INPUT
	ECLASSID : DINT;
END_VAR
END_METHOD

METHOD OCCUPYRESOURCE : BOOL
VAR_INPUT
	ECLASSID : DINT;
END_VAR
END_METHOD

METHOD SETCAPACITY
VAR_INPUT
	ITFLISTCONTROL : L_UBUP_IListControl;
	DWCAPACITY : DWORD;
END_VAR
END_METHOD

METHOD SETCAPACITYALL
END_METHOD

METHOD FB_INIT : BOOL
VAR_INPUT
	BINITRETAINS : BOOL;
	BINCOPYCODE : BOOL;
	PICKANDPLACEMEMORY : REFERENCE TO L_MC4P_PickAndPlaceMemory;
	SCFBSTORE : REFERENCE TO L_MC4P_MovePathStore;
END_VAR
END_METHOD

METHOD FREERESOURCE
END_METHOD

METHOD GETFB : L_UBUP_IPoolInstance
VAR_INPUT
	ECLASSID : DINT;
	DWARRIDX : DWORD;
END_VAR
END_METHOD

METHOD GETFBCONTROL : L_UBUP_IListControl
VAR_INPUT
	ECLASSID : DINT;
END_VAR
END_METHOD

METHOD OCCUPYRESOURCE : BOOL
VAR_INPUT
	ECLASSID : DINT;
END_VAR
END_METHOD

METHOD SETCAPACITYALL
END_METHOD

(* ---- L_MC4P_MOVELINEARABSOLUTE_INTERNAL.fb ---- *)
FUNCTION_BLOCK L_MC4P_MOVELINEARABSOLUTE_INTERNAL EXTENDS L_MC4P_MoveContPath
VAR_INPUT
	EXECUTE : BOOL;
	POSITION : ARRAY [1..12] OF LREAL;
	VELOCITY : LREAL;
	ACCELERATION : LREAL;
	DECELERATION : LREAL;
	JERK : LREAL;
	COORDSYSTEM : L_MC4P_CoordSystem;
	BUFFERMODE : MC_BUFFER_MODE;
	TRANSITIONMODE : MC_TRANSITION_MODE;
	TRANSITIONPARAMETER : ARRAY [1..12] OF LREAL := [12(0)];
	AEAUXMODE : ARRAY [1..6] OF L_MC4P_AuxMode;
	ORIENTATIONMODE : L_MC4P_Orientation_Mode := L_MC4P_Orientation_Mode.ShortestSpacialWay;
	DIRECTION : ARRAY [4..6] OF MC_DIRECTION := [3(MC_DIRECTION.mcShortestWay)];
END_VAR
VAR_OUTPUT
	DONE : BOOL;
	BUSY : BOOL;
	ACTIVE : BOOL;
	COMMANDABORTED : BOOL;
	ERROR : BOOL;
	ERRORID : L_IE1P_Error;
END_VAR
VAR
	CLASSID : DINT;
END_VAR
END_FUNCTION_BLOCK

METHOD HOMINGREQUIRED : BOOL
END_METHOD

METHOD MAIN
VAR_IN_OUT
	AXESGROUP : AXES_GROUP_KIN;
	FBBASE : L_MC4P_Template_AG_KIN;
END_VAR
END_METHOD

METHOD PARAMETERFREEZE
VAR_IN_OUT
	AXESGROUP : AXES_GROUP_KIN;
	FBBASE : L_MC4P_Template_AG_KIN;
	COORDSYSTEM : L_MC4P_CoordSystem;
	BUFFERMODE : MC_BUFFER_MODE;
	TRANSITIONMODE : MC_TRANSITION_MODE;
	TRANSITIONPARAMETER : ARRAY [1..12] OF LREAL;
END_VAR
END_METHOD

METHOD SETERRORINPUTLIMITATIONVIOLATION
VAR_IN_OUT
	FBBASE : L_MC4P_Template_AG_KIN;
END_VAR
END_METHOD

METHOD SETPATHELEMENT
VAR_IN_OUT
	AXESGROUP : AXES_GROUP_KIN;
	FBBASE : L_MC4P_Template_AG_KIN;
	ALRSTARTPOS : ARRAY [1..12] OF LREAL;
	ALRSUPERPOSPOSATSTART : ARRAY [1..3] OF LREAL;
END_VAR
END_METHOD

(* ---- L_MC4P_MOVELINEARRELATIVE_INTERNAL.fb ---- *)
FUNCTION_BLOCK L_MC4P_MOVELINEARRELATIVE_INTERNAL EXTENDS L_MC4P_MoveContPath
VAR_INPUT
	EXECUTE : BOOL;
	DISTANCE : ARRAY [1..12] OF LREAL;
	VELOCITY : LREAL;
	ACCELERATION : LREAL;
	DECELERATION : LREAL;
	JERK : LREAL;
	COORDSYSTEM : L_MC4P_CoordSystem;
	BUFFERMODE : MC_BUFFER_MODE;
	TRANSITIONMODE : MC_TRANSITION_MODE;
	TRANSITIONPARAMETER : ARRAY [1..12] OF LREAL := [12(0)];
	AEAUXMODE : ARRAY [1..6] OF L_MC4P_AuxMode;
	ORIENTATIONMODE : L_MC4P_Orientation_Mode := L_MC4P_Orientation_Mode.ShortestSpacialWay;
	DIRECTION : ARRAY [4..6] OF MC_DIRECTION := [3(MC_DIRECTION.mcShortestWay)];
END_VAR
VAR_OUTPUT
	DONE : BOOL;
	BUSY : BOOL;
	ACTIVE : BOOL;
	COMMANDABORTED : BOOL;
	ERROR : BOOL;
	ERRORID : L_IE1P_Error;
END_VAR
VAR
	CLASSID : DINT;
END_VAR
END_FUNCTION_BLOCK

METHOD HOMINGREQUIRED : BOOL
END_METHOD

METHOD MAIN
VAR_IN_OUT
	AXESGROUP : AXES_GROUP_KIN;
	FBBASE : L_MC4P_Template_AG_KIN;
END_VAR
END_METHOD

METHOD PARAMETERFREEZE
VAR_IN_OUT
	AXESGROUP : AXES_GROUP_KIN;
	FBBASE : L_MC4P_Template_AG_KIN;
	COORDSYSTEM : L_MC4P_CoordSystem;
	BUFFERMODE : MC_BUFFER_MODE;
	TRANSITIONMODE : MC_TRANSITION_MODE;
	TRANSITIONPARAMETER : ARRAY [1..12] OF LREAL;
END_VAR
END_METHOD

METHOD SETERRORINPUTLIMITATIONVIOLATION
VAR_IN_OUT
	FBBASE : L_MC4P_Template_AG_KIN;
END_VAR
END_METHOD

METHOD SETPATHELEMENT
VAR_IN_OUT
	AXESGROUP : AXES_GROUP_KIN;
	FBBASE : L_MC4P_Template_AG_KIN;
	ALRSTARTPOS : ARRAY [1..12] OF LREAL;
	ALRSUPERPOSPOSATSTART : ARRAY [1..3] OF LREAL;
END_VAR
END_METHOD

(* ---- L_MC4P_MOVESPLINEABSOLUTE.fb ---- *)
FUNCTION_BLOCK L_MC4P_MOVESPLINEABSOLUTE EXTENDS L_MC4P_Template_MoveLicence
VAR_INPUT
	XEXECUTE : BOOL;
	ASCINTERMEDIATEPOINT : ARRAY [1..9] OF L_MC4P_IntermediatePointSpline;
	ALRENDPOINT : ARRAY [1..12] OF LREAL;
	LRVELOCITY : LREAL;
	LRACCELERATION : LREAL;
	LRDECELERATION : LREAL;
	LRJERK : LREAL;
	ECOORDSYSTEM : L_MC4P_CoordSystem;
	EBUFFERMODE : MC_BUFFER_MODE;
	ETRANSITIONMODE : MC_TRANSITION_MODE;
	ALRTRANSITIONPARAMETER : ARRAY [1..12] OF LREAL := [12(0)];
	AEAUXMODE : ARRAY [1..6] OF L_MC4P_AuxMode;
	EORIENTATIONMODE : L_MC4P_Orientation_Mode := L_MC4P_Orientation_Mode.ShortestSpacialWay;
	AEDIRECTION : ARRAY [4..6] OF MC_DIRECTION := [3(MC_DIRECTION.mcShortestWay)];
END_VAR
VAR_OUTPUT
	XDONE : BOOL;
	XBUSY : BOOL;
	XACTIVE : BOOL;
	XCOMMANDABORTED : BOOL;
	XERROR : BOOL;
	EERRORID : L_IE1P_Error;
	IPOINTPASSED : INT;
END_VAR
VAR
	MOVESPLINE : L_MC4P_MoveSplineAbsolute_Internal;
	XDIALOGINTERMEDIATEPOINT : BOOL := FALSE;
	IVISUTABLESETPOS : INT := 1;
	PASSEDINTERMEDIATEPOINT : INT;
	PMOVE : POINTER TO L_MC4P_MoveContPath;
END_VAR
END_FUNCTION_BLOCK

(* ---- L_MC4P_MOVESPLINEABSOLUTE_INTERNAL.fb ---- *)
FUNCTION_BLOCK L_MC4P_MOVESPLINEABSOLUTE_INTERNAL EXTENDS L_MC4P_MoveContPath
VAR_INPUT
	XEXECUTE : BOOL;
	ASCINTERMEDIATEPOINT : ARRAY [1..9] OF L_MC4P_IntermediatePointSpline;
	ALRENDPOINT : ARRAY [1..12] OF LREAL;
	LRVELOCITY : LREAL;
	LRACCELERATION : LREAL;
	LRDECELERATION : LREAL;
	LRJERK : LREAL;
	ECOORDSYSTEM : L_MC4P_CoordSystem;
	EBUFFERMODE : MC_BUFFER_MODE;
	ETRANSITIONMODE : MC_TRANSITION_MODE;
	ALRTRANSITIONPARAMETER : ARRAY [1..12] OF LREAL := [12(0)];
	AEAUXMODE : ARRAY [1..6] OF L_MC4P_AuxMode;
	EORIENTATIONMODE : L_MC4P_Orientation_Mode := L_MC4P_Orientation_Mode.ShortestSpacialWay;
	AEDIRECTION : ARRAY [4..6] OF MC_DIRECTION := [3(MC_DIRECTION.mcShortestWay)];
END_VAR
VAR_OUTPUT
	XDONE : BOOL;
	XBUSY : BOOL;
	XACTIVE : BOOL;
	XCOMMANDABORTED : BOOL;
	XERROR : BOOL;
	EERRORID : L_IE1P_Error;
	IPOINTPASSED : INT;
END_VAR
VAR
	CLASSID : DINT;
	PASSEDINTERMEDIATEPOINT : INT;
END_VAR
END_FUNCTION_BLOCK

METHOD HOMINGREQUIRED : BOOL
END_METHOD

METHOD MAIN
VAR_IN_OUT
	AXESGROUP : AXES_GROUP_KIN;
	FBBASE : L_MC4P_Template_AG_KIN;
END_VAR
END_METHOD

METHOD PARAMETERFREEZE
VAR_IN_OUT
	AXESGROUP : AXES_GROUP_KIN;
	FBBASE : L_MC4P_Template_AG_KIN;
	COORDSYSTEM : L_MC4P_CoordSystem;
	BUFFERMODE : MC_BUFFER_MODE;
	TRANSITIONMODE : MC_TRANSITION_MODE;
	TRANSITIONPARAMETER : ARRAY [1..12] OF LREAL;
END_VAR
END_METHOD

METHOD SETERRORINPUTLIMITATIONVIOLATION
VAR_IN_OUT
	FBBASE : L_MC4P_Template_AG_KIN;
END_VAR
END_METHOD

METHOD SETPATHELEMENT
VAR_IN_OUT
	AXESGROUP : AXES_GROUP_KIN;
	FBBASE : L_MC4P_Template_AG_KIN;
	ALRSTARTPOS : ARRAY [1..12] OF LREAL;
	ALRSUPERPOSPOSATSTART : ARRAY [1..3] OF LREAL;
END_VAR
END_METHOD

(* ---- L_MC4P_MOVESPLINEPNP.fb ---- *)
FUNCTION_BLOCK L_MC4P_MOVESPLINEPNP EXTENDS L_MC4P_Template_MoveLicence
VAR_INPUT
	XEXECUTE : BOOL;
	LRZSTARTDIST : LREAL;
	LRZTARGETDIST : LREAL;
	ALRENDPOINT : ARRAY [1..12] OF LREAL;
	LRZMAXHEIGHT : LREAL;
	LRVELOCITY : LREAL;
	LRACCELERATION : LREAL;
	LRDECELERATION : LREAL;
	LRJERK : LREAL;
	ECOORDSYSTEM : L_MC4P_CoordSystem;
	EBUFFERMODE : MC_BUFFER_MODE;
	ETRANSITIONMODE : MC_TRANSITION_MODE;
	ALRTRANSITIONPARAMETER : ARRAY [1..12] OF LREAL := [12(0)];
	AEAUXMODE : ARRAY [1..6] OF L_MC4P_AuxMode;
	EORIENTATIONMODE : L_MC4P_Orientation_Mode := L_MC4P_Orientation_Mode.ShortestSpacialWay;
	AEDIRECTION : ARRAY [4..6] OF MC_DIRECTION := [3(MC_DIRECTION.mcShortestWay)];
END_VAR
VAR_OUTPUT
	XDONE : BOOL;
	XBUSY : BOOL;
	XACTIVE : BOOL;
	XCOMMANDABORTED : BOOL;
	XERROR : BOOL;
	EERRORID : L_IE1P_Error;
	IPOINTPASSED : INT;
END_VAR
VAR
	MOVESPLINE : L_MC4P_MoveSplinePnP_Internal;
	PASSEDINTERMEDIATEPOINT : INT;
	PMOVE : POINTER TO L_MC4P_MoveContPath;
END_VAR
END_FUNCTION_BLOCK

(* ---- L_MC4P_MOVESPLINEPNP_INTERNAL.fb ---- *)
FUNCTION_BLOCK L_MC4P_MOVESPLINEPNP_INTERNAL EXTENDS L_MC4P_MoveContPath
VAR_INPUT
	XEXECUTE : BOOL;
	LRZSTARTDIST : LREAL;
	LRZTARGETDIST : LREAL;
	ALRENDPOINT : ARRAY [1..12] OF LREAL;
	LRZMAXHEIGHT : LREAL;
	LRVELOCITY : LREAL;
	LRACCELERATION : LREAL;
	LRDECELERATION : LREAL;
	LRJERK : LREAL;
	ECOORDSYSTEM : L_MC4P_CoordSystem;
	EBUFFERMODE : MC_BUFFER_MODE;
	ETRANSITIONMODE : MC_TRANSITION_MODE;
	ALRTRANSITIONPARAMETER : ARRAY [1..12] OF LREAL := [12(0)];
	AEAUXMODE : ARRAY [1..6] OF L_MC4P_AuxMode;
	EORIENTATIONMODE : L_MC4P_Orientation_Mode := L_MC4P_Orientation_Mode.ShortestSpacialWay;
	AEDIRECTION : ARRAY [4..6] OF MC_DIRECTION := [3(MC_DIRECTION.mcShortestWay)];
END_VAR
VAR_OUTPUT
	XDONE : BOOL;
	XBUSY : BOOL;
	XACTIVE : BOOL;
	XCOMMANDABORTED : BOOL;
	XERROR : BOOL;
	EERRORID : L_IE1P_Error;
	IPOINTPASSED : INT;
END_VAR
VAR
	CLASSID : DINT;
	PASSEDINTERMEDIATEPOINT : INT;
END_VAR
END_FUNCTION_BLOCK

METHOD HOMINGREQUIRED : BOOL
END_METHOD

METHOD MAIN
VAR_IN_OUT
	AXESGROUP : AXES_GROUP_KIN;
	FBBASE : L_MC4P_Template_AG_KIN;
END_VAR
END_METHOD

METHOD PARAMETERFREEZE
VAR_IN_OUT
	AXESGROUP : AXES_GROUP_KIN;
	FBBASE : L_MC4P_Template_AG_KIN;
	COORDSYSTEM : L_MC4P_CoordSystem;
	BUFFERMODE : MC_BUFFER_MODE;
	TRANSITIONMODE : MC_TRANSITION_MODE;
	TRANSITIONPARAMETER : ARRAY [1..12] OF LREAL;
END_VAR
END_METHOD

METHOD SETERRORINPUTLIMITATIONVIOLATION
VAR_IN_OUT
	FBBASE : L_MC4P_Template_AG_KIN;
END_VAR
END_METHOD

METHOD SETPATHELEMENT
VAR_IN_OUT
	AXESGROUP : AXES_GROUP_KIN;
	FBBASE : L_MC4P_Template_AG_KIN;
	ALRSTARTPOS : ARRAY [1..12] OF LREAL;
	ALRSUPERPOSPOSATSTART : ARRAY [1..3] OF LREAL;
END_VAR
END_METHOD

(* ---- L_MC4P_MOVESPLINERELATIVE.fb ---- *)
FUNCTION_BLOCK L_MC4P_MOVESPLINERELATIVE EXTENDS L_MC4P_Template_MoveLicence
VAR_INPUT
	XEXECUTE : BOOL;
	ASCINTERMEDIATEPOINT : ARRAY [1..9] OF L_MC4P_IntermediatePointSpline;
	ALRENDPOINT : ARRAY [1..12] OF LREAL;
	LRVELOCITY : LREAL;
	LRACCELERATION : LREAL;
	LRDECELERATION : LREAL;
	LRJERK : LREAL;
	ECOORDSYSTEM : L_MC4P_CoordSystem;
	EBUFFERMODE : MC_BUFFER_MODE;
	ETRANSITIONMODE : MC_TRANSITION_MODE;
	ALRTRANSITIONPARAMETER : ARRAY [1..12] OF LREAL := [12(0)];
	AEAUXMODE : ARRAY [1..6] OF L_MC4P_AuxMode;
	EORIENTATIONMODE : L_MC4P_Orientation_Mode := L_MC4P_Orientation_Mode.ShortestSpacialWay;
	AEDIRECTION : ARRAY [4..6] OF MC_DIRECTION := [3(MC_DIRECTION.mcShortestWay)];
END_VAR
VAR_OUTPUT
	XDONE : BOOL;
	XBUSY : BOOL;
	XACTIVE : BOOL;
	XCOMMANDABORTED : BOOL;
	XERROR : BOOL;
	EERRORID : L_IE1P_Error;
	IPOINTPASSED : INT;
END_VAR
VAR
	MOVESPLINE : L_MC4P_MoveSplineRelative_Internal;
	XDIALOGINTERMEDIATEPOINT : BOOL := FALSE;
	IVISUTABLESETPOS : INT := 1;
	PASSEDINTERMEDIATEPOINT : INT;
	PMOVE : POINTER TO L_MC4P_MoveContPath;
END_VAR
END_FUNCTION_BLOCK

(* ---- L_MC4P_MOVESPLINERELATIVE_INTERNAL.fb ---- *)
FUNCTION_BLOCK L_MC4P_MOVESPLINERELATIVE_INTERNAL EXTENDS L_MC4P_MoveContPath
VAR_INPUT
	XEXECUTE : BOOL;
	ASCINTERMEDIATEPOINT : ARRAY [1..9] OF L_MC4P_IntermediatePointSpline;
	ALRENDPOINT : ARRAY [1..12] OF LREAL;
	LRVELOCITY : LREAL;
	LRACCELERATION : LREAL;
	LRDECELERATION : LREAL;
	LRJERK : LREAL;
	ECOORDSYSTEM : L_MC4P_CoordSystem;
	EBUFFERMODE : MC_BUFFER_MODE;
	ETRANSITIONMODE : MC_TRANSITION_MODE;
	ALRTRANSITIONPARAMETER : ARRAY [1..12] OF LREAL := [12(0)];
	AEAUXMODE : ARRAY [1..6] OF L_MC4P_AuxMode;
	EORIENTATIONMODE : L_MC4P_Orientation_Mode := L_MC4P_Orientation_Mode.ShortestSpacialWay;
	AEDIRECTION : ARRAY [4..6] OF MC_DIRECTION := [3(MC_DIRECTION.mcShortestWay)];
END_VAR
VAR_OUTPUT
	XDONE : BOOL;
	XBUSY : BOOL;
	XACTIVE : BOOL;
	XCOMMANDABORTED : BOOL;
	XERROR : BOOL;
	EERRORID : L_IE1P_Error;
	IPOINTPASSED : INT;
END_VAR
VAR
	CLASSID : DINT;
	PASSEDINTERMEDIATEPOINT : INT;
END_VAR
END_FUNCTION_BLOCK

METHOD HOMINGREQUIRED : BOOL
END_METHOD

METHOD MAIN
VAR_IN_OUT
	AXESGROUP : AXES_GROUP_KIN;
	FBBASE : L_MC4P_Template_AG_KIN;
END_VAR
END_METHOD

METHOD PARAMETERFREEZE
VAR_IN_OUT
	AXESGROUP : AXES_GROUP_KIN;
	FBBASE : L_MC4P_Template_AG_KIN;
	COORDSYSTEM : L_MC4P_CoordSystem;
	BUFFERMODE : MC_BUFFER_MODE;
	TRANSITIONMODE : MC_TRANSITION_MODE;
	TRANSITIONPARAMETER : ARRAY [1..12] OF LREAL;
END_VAR
END_METHOD

METHOD SETERRORINPUTLIMITATIONVIOLATION
VAR_IN_OUT
	FBBASE : L_MC4P_Template_AG_KIN;
END_VAR
END_METHOD

METHOD SETPATHELEMENT
VAR_IN_OUT
	AXESGROUP : AXES_GROUP_KIN;
	FBBASE : L_MC4P_Template_AG_KIN;
	ALRSTARTPOS : ARRAY [1..12] OF LREAL;
	ALRSUPERPOSPOSATSTART : ARRAY [1..3] OF LREAL;
END_VAR
END_METHOD

(* ---- L_MC4P_OBSERVELIMITS.fb ---- *)
FUNCTION_BLOCK L_MC4P_OBSERVELIMITS
VAR_INPUT
	XENABLE : BOOL;
	XRESETOBSERVEDLIMITS : BOOL;
	XHOLDOBSERVEDLIMITS : BOOL;
	PAXESGROUP : POINTER TO AXES_GROUP_KIN;
	UACTIVELIMITSMAN : L_MC1P.L_MC1P_uULINT;
END_VAR
VAR_OUTPUT
	UACTIVELIMITS : L_MC1P.L_MC1P_uULINT;
END_VAR
VAR
	XENABLEOLD : BOOL;
	IDX : INT;
	PAXIS : POINTER TO AXIS_REF;
	ALRSETACCOLD : ARRAY [1..6] OF LREAL;
	ALRSETJERK : ARRAY [1..6] OF LREAL;
	LRMAXVELFB : LREAL;
	LRMAXACCFB : LREAL;
	LRMAXJERKFB : LREAL;
	SCLAMPACTIVAX : ARRAY [1..12, 1..10, 0..1] OF BOOL;
	SCLAMPACTIVAG : ARRAY [1..3, 1..3, 0..1] OF BOOL;
	WVISUAXESFRAME : WORD;
	HEVENTCOMMCYCLE : Systypes.RTS_IEC_HANDLE := SysTypes.RTS_INVALID_HANDLE;
	HINTERFACECOMMCYCLE : Systypes.RTS_IEC_HANDLE := SysTypes.RTS_INVALID_HANDLE;
	ITFCALLBACK : CmpEventMgr.ICmpEventCallback;
	DWEVENTCOUNTER : DWORD;
END_VAR
END_FUNCTION_BLOCK

METHOD LIMITUSED : BOOL
VAR_INPUT
	LRCMPVAL : LREAL;
	LRACTVAL : LREAL;
END_VAR
END_METHOD

METHOD MAIN
END_METHOD

METHOD SETLAMPACTIV
END_METHOD

METHOD EVENTCALLBACK : UDINT
VAR_INPUT
	PEVENTPARAM : POINTER TO EventParam;
END_VAR
END_METHOD

METHOD REGISTEREVENT
END_METHOD

METHOD UNREGISTEREVENT
END_METHOD

(* ---- L_MC4P_PATHDATALIST.fb ---- *)
FUNCTION_BLOCK L_MC4P_PATHDATALIST
VAR_INPUT
	PAXESGROUP : POINTER TO AXES_GROUP_KIN;
END_VAR
VAR
	PLISTELEMENTFIRST : POINTER TO L_MC4P_ListElement;
	PLISTELEMENTLAST : POINTER TO L_MC4P_ListElement;
	XINITDONE : BOOL := FALSE;
	ARRLISTELEMENTS : ARRAY [0..L_MC4P_Constants.MaxCountListElements] OF L_MC4P_ListElement;
	SCINITIALLISTELEMENT : L_MC4P_ListElement;
END_VAR
END_FUNCTION_BLOCK

METHOD CALCPATHLENGTHLISTELEMENTS : LREAL
VAR_INPUT
	DWMASK : DWORD;
END_VAR
END_METHOD

METHOD CALCPATHLENGTHLISTELEMENTSOFFUNID : LREAL
VAR_INPUT
	DIFUNID : DINT;
END_VAR
END_METHOD

METHOD CALCTIMELISTELEMENTS : LREAL
VAR_INPUT
	DWMASK : DWORD;
END_VAR
END_METHOD

METHOD CALCTIMELISTELEMENTSOFFUNID : LREAL
VAR_INPUT
	DIFUNID : DINT;
END_VAR
END_METHOD

METHOD CHECKLIST : BOOL
END_METHOD

METHOD CHECKLISTANDPROFILES : BOOL
END_METHOD

METHOD CLEARFBPOINTER
VAR_INPUT
	PMOVECONTFB : POINTER TO L_MC4P_MoveContPath;
END_VAR
END_METHOD

METHOD COUNTLISTELEMENTS : INT
VAR_INPUT
	DWMASK : DWORD;
END_VAR
END_METHOD

METHOD DELETELISTELEMENT : BOOL
VAR_INPUT
	PLISTELEMENT : POINTER TO L_MC4P_ListElement;
END_VAR
END_METHOD

METHOD GETLISTELEMENTBYTIME : POINTER TO L_MC4P_ListElement
VAR_INPUT
	DWMASK : DWORD;
	LRTIMELISTIN : LREAL;
END_VAR
VAR_OUTPUT
	LRTIMEELEMENT : LREAL;
END_VAR
END_METHOD

METHOD GETLISTELEMENTOFFUNID : POINTER TO L_MC4P_ListElement
VAR_INPUT
	DIFUNID : DINT;
END_VAR
END_METHOD

METHOD GETNEWESTLISTELEMENT : POINTER TO L_MC4P_ListElement
VAR_INPUT
	DWMASK : DWORD;
END_VAR
END_METHOD

METHOD GETOLDESTLISTELEMENT : POINTER TO L_MC4P_ListElement
VAR_INPUT
	DWMASK : DWORD;
END_VAR
END_METHOD

METHOD GETOLDESTLISTELEMENTADVANCED : POINTER TO L_MC4P_ListElement
VAR_INPUT
	DWMASK : DWORD;
	DWPREVMASK : DWORD;
END_VAR
END_METHOD

METHOD INITLIST : BOOL
END_METHOD

METHOD INITLISTELEMENT : BOOL
VAR_INPUT
	PLISTELEMENT : POINTER TO L_MC4P_ListElement;
END_VAR
END_METHOD

METHOD INSERTLISTELEMENTBETWEEN : POINTER TO L_MC4P_ListElement
VAR_INPUT
	PPREVIOUS : POINTER TO L_MC4P_ListElement;
END_VAR
END_METHOD

METHOD INSERTNEWLISTELEMENT : POINTER TO L_MC4P_ListElement
END_METHOD

METHOD NUMLISTELEMENTSISLESSTHAN : BOOL
VAR_INPUT
	DWMASK : DWORD;
	IUPPER : INT;
END_VAR
END_METHOD

METHOD RESETLIST
END_METHOD

METHOD RESETMASKSINLIST
VAR_INPUT
	FIPOSECTIME : LREAL;
END_VAR
END_METHOD

METHOD STARTVELOFLISTELEMENTEQ0 : BOOL
VAR_INPUT
	PLISTELEMENT : POINTER TO L_MC4P_ListElement;
END_VAR
END_METHOD

METHOD TARGETVELOFLISTELEMENTEQ0 : BOOL
VAR_INPUT
	PLISTELEMENT : POINTER TO L_MC4P_ListElement;
END_VAR
END_METHOD

METHOD TIMELISTELEMENTSISLESSTHAN : BOOL
VAR_INPUT
	DWMASK : DWORD;
	LRUPPER : LREAL;
END_VAR
END_METHOD

METHOD _CREATELISTELEMENT : POINTER TO L_MC4P_ListElement
END_METHOD

METHOD _DESTROYLISTELEMENT
VAR_INPUT
	PLISTELEMENT : POINTER TO L_MC4P_ListElement;
END_VAR
END_METHOD

(* ---- L_MC4P_PATHLISTDIAGNOSTIC.fb ---- *)
FUNCTION_BLOCK L_MC4P_PATHLISTDIAGNOSTIC
VAR_INPUT
	XWRITEFILEEXECUTE : BOOL;
	XREADERRORFILEEXECUTE : BOOL;
	XENABLE : BOOL;
	INUMOFLISTELEMENTS : INT;
END_VAR
VAR_OUTPUT
	XWRITEFILEDONE : BOOL;
	XWRITEFILEBUSY : BOOL;
	XWRITEFILEERROR : BOOL;
	XERRORDETECTED : BOOL;
	XCHECKCONSISTENCYFAIL : BOOL;
	XDONE : BOOL;
	XBUSY : BOOL;
	AL_MC4P_LISTELEMENT : ARRAY [0..(ciArrayBreite + ciArrayHistory)] OF L_MC4P_ListElement;
	INUMOFLISTELEMENTSOUT : INT;
	APLISTELEM : ARRAY [0..(ciArrayBreite + ciArrayHistory)] OF POINTER TO L_MC4P_ListElement;
	ILISTHISTORYEND : INT := 1;
	ASCLISTHISTORY : ARRAY [1..ciArrayHistory] OF L_MC4P_ListElement;
END_VAR
VAR
	CIARRAYHISTORY : INT := 10;
	CIARRAYTIEFE : INT := 1000;
	CIARRAYBREITE : INT := 30;
	XTESTINMOTIONTASK : BOOL := FALSE;
	XFREETASKBUSY_INT : BOOL;
	XFREETASKDONE_INT : BOOL;
	XFREETASKERROR_INT : BOOL;
	EFREETASKEERRORID_INT : L_IE1P_Error;
	RES : SYSFILE.RTS_IEC_ResULT;
	HFILE : SYSFILE.RTS_IEC_HANDLE;
	XWFSIZE : __XWORD;
	XWRESULTWRITESTRING : __XWORD;
	FB_STACKDIAGDATA : L_MC1P_StackControlArray := STRUCT(iMaxLegth := ciArrayTiefe);
	ASCDIAGDATA : ARRAY [0..ciArrayTiefe] OF L_MC4P_PathListDiagnosticData;
	SCDIAGDATATMP : L_MC4P_PathListDiagnosticData;
	WSTEP : WORD := 0;
	WSTEPREF : WORD := 0;
	WSTEPWEF : WORD := 0;
	WSTEPWF : WORD := 0;
	XDATACHENGED : BOOL;
	XCONSISTENCY : BOOL;
	XWRITEFILEEXECUTE_OLD : BOOL;
	IDX : INT;
	INUMOFLISTELEMENTS_INT : INT;
	PLISTELEMENTLAST : POINTER TO L_MC4P_ListElement;
	PLISTELEMENTFIRST : POINTER TO L_MC4P_ListElement;
	PLEFT : POINTER TO L_MC4P_ListElement;
	OPEN2 : FILE.Open;
	CLOSE2 : FILE.Close;
	READ1 : FILE.Read;
	ASHEADLINE : ARRAY [1..10] OF STRING(255) := ['Hinweise zur ListenElementen:  Segmentnummer +2000:  Element aus Ipo,  Segmentnummer +1000:  diSegmentNoCopiedFrom $N', 'Hinweise zur Exeltabelle: oben ist der älteste und unten ist der akttuelste Stand der Liste  $N', 'Zeile1:AnzahlDurchläufe $TxPathStopExecute $TdiActFunID $TdiBusyFunID $TdiFunID $TlrOverride $T $TSegmente  $N', 'Zeile2: AbsZähler $TxPathStopExecute $TdiActFunID $TdiBusyFunID $TdiFunID, $TlrOverride $T $TMaske $T $N', '$N '];
	STABULATOR : STRING(2) := '$T';
	SLINEFEED : STRING(2) := '$N';
	SZEILE : STRING(255);
	SZEILE2 : STRING(255);
	IDATAIDX1 : INT;
	SEXELFILENAME : STRING;
	SLISTELEMENTFILENAME : STRING;
	SLISTELEMENTFILENAMEBASE : STRING;
	XREADERRORFILEDONE : BOOL;
	XREADERRORFILEBUSY : BOOL;
	XREADERRORFILEERROR : BOOL;
	XWRITEFILEEXECUTE_INTERN : BOOL;
	XREADERRORFILEEXECUTE_INTERN : BOOL;
	XREADERRORFILEEXECUTE_OLD : BOOL;
	DITIMESTAMP : DINT;
	ILISTHISTORYENDLENGTH : INT;
	SCLISTELEMENTEMPTY : L_MC4P_ListElement;
	IDX2 : INT;
	IDX3 : INT;
	ILISTELEMACTIVE : INT;
	IDATANO : INT;
	XAGERORR : BOOL;
	ASCAGEERRORINFO : ARRAY [0..7] OF L_IE1P_ErrorInformation;
	XSAVEAGERROR : BOOL;
	WLOOKAHEADHORIZON : WORD;
	DWTASKYCLE_US : DWORD;
	EACTIVEERRORID : L_IE1P_Error;
	SAXESGROUPNAME : STRING;
	XWRITEINMOTIONTASK : BOOL;
END_VAR
END_FUNCTION_BLOCK

METHOD CALL_CHECKCHANGES_SCDIAGDATA : BOOL
VAR_IN_OUT
	SCDIAGDATANEW : L_MC4P_PathListDiagnosticData;
	SCDIAGDATAOLD : L_MC4P_PathListDiagnosticData;
END_VAR
END_METHOD

METHOD CALL_CHECKCONSISTENCY : BOOL
VAR_IN_OUT
	SCDIAGDATA : L_MC4P_PathListDiagnosticData;
END_VAR
END_METHOD

METHOD CALL_INIT_SCDIAGDATA
VAR_IN_OUT
	SCDIAGDATA : L_MC4P_PathListDiagnosticData;
END_VAR
END_METHOD

METHOD CHECKCONSISTENCY
END_METHOD

METHOD READERRORFILE
END_METHOD

METHOD MAINFB : BOOL
VAR_INPUT
	PAXESGROUP : POINTER TO AXES_GROUP_KIN;
END_VAR
END_METHOD

METHOD CALL_WRITEEXELFILE
END_METHOD

METHOD CALL_WRITESEGEMENTFILE
VAR_IN_OUT
	SCLISTELEM : L_MC4P_ListElement;
END_VAR
END_METHOD

METHOD EXECUTEFREERUNTASK
END_METHOD

METHOD MAIN
END_METHOD

METHOD RESETREADDATA
END_METHOD

METHOD ABORT : UDINT
END_METHOD

METHOD EXECUTE : UDINT
END_METHOD
